FUNCTION "ROLL_PB13" : Void
{ S7_Optimized_Access := 'TRUE' }
VERSION : 0.1
VAR_TEMP
    r : Bool;
    a1 : Word;
    a2 : Word;
    activeDataBlock : Int;
    comparisonResults : Array[0..0] of Bool;
END_VAR
BEGIN
    #r := FALSE;
    #a1 := W#16#0000;
    #a2 := W#16#0000;
    #activeDataBlock := 0;
    // PB13, STEP 5 network 1
    #r := ((NOT "ROLL_State".M[58, 6]) AND ("ROLL_IO".Input[11, 1] OR "ROLL_IO".Input[11, 2] OR "ROLL_IO".Input[11, 3] OR "ROLL_IO".Input[11, 4] OR "ROLL_IO".Input[119, 6] OR "ROLL_IO".Input[119, 7] OR "ROLL_IO".Input[120, 0]) AND "ROLL_IO".Input[11, 6]);
    IF #r THEN "ROLL_State".M[58, 7] := TRUE; END_IF;
    #r := (((NOT "ROLL_IO".Input[11, 6]) AND ("ROLL_IO".Input[11, 1] OR "ROLL_IO".Input[11, 2] OR "ROLL_IO".Input[11, 3] OR "ROLL_IO".Input[11, 4] OR "ROLL_IO".Input[119, 6] OR "ROLL_IO".Input[119, 7] OR "ROLL_IO".Input[120, 0]) AND "ROLL_IO".Output[23, 0] AND "ROLL_State".M[58, 6]) OR "ROLL_IO".Input[11, 0]);
    IF #r THEN "ROLL_State".M[58, 7] := FALSE; END_IF;
    // PB13, STEP 5 network 2
    #r := "ROLL_IO".Input[11, 6];
    "ROLL_State".M[58, 6] := #r;
    // PB13, STEP 5 network 3
    #r := (((((NOT "ROLL_IO".Input[11, 0]) OR "ROLL_State".M[80, 7]) AND "ROLL_IO".Input[11, 6]) OR "ROLL_State".M[58, 7]) AND "ROLL_IO".Input[14, 0]);
    "ROLL_State".M[60, 0] := #r;
    // PB13, STEP 5 network 4
    #a2 := #a1;
    #a1 := W#16#2030;
    #r := ((NOT "ROLL_IO".Input[13, 3]) AND "ROLL_IO".Output[24, 0]);
    "ROLL_TimerOp"(Number := 110, Operation := 0, Signal := #r, Preset := #a1);
    // PB13, STEP 5 network 5
    #r := (((NOT "ROLL_State".M[111, 1]) AND (NOT "ROLL_State".M[111, 2]) AND (NOT "ROLL_State".M[111, 5]) AND "ROLL_IO".Input[0, 2] AND "ROLL_State".M[111, 0]) OR ((NOT "ROLL_State".M[61, 5]) AND "ROLL_IO".Input[0, 1] AND "ROLL_State".M[23, 2]) OR ("ROLL_IO".Input[12, 1] AND "ROLL_State".M[111, 5]));
    "ROLL_State".M[60, 1] := #r;
    // PB13, STEP 5 network 6
    #r := (((NOT "ROLL_IO".Input[12, 1]) AND "ROLL_State".M[111, 5]) OR ((NOT "ROLL_State".M[111, 0]) AND (NOT "ROLL_State".M[111, 2]) AND (NOT "ROLL_State".M[111, 5]) AND "ROLL_IO".Input[0, 2] AND "ROLL_State".M[111, 1]) OR ("ROLL_IO".Input[0, 1] AND "ROLL_State".M[23, 3]));
    "ROLL_State".M[60, 3] := #r;
    // PB13, STEP 5 network 7
    #r := (((NOT "ROLL_State".M[111, 0]) AND (NOT "ROLL_State".M[111, 1]) AND (NOT "ROLL_State".M[111, 5]) AND "ROLL_IO".Input[0, 2] AND "ROLL_State".M[111, 2]) OR ((NOT "ROLL_State".M[61, 5]) AND "ROLL_IO".Input[0, 1] AND "ROLL_State".M[0, 3]));
    "ROLL_State".M[60, 2] := #r;
    // PB13, STEP 5 network 8
    #a2 := #a1;
    #a1 := W#16#0005;
    #r := (NOT "ROLL_State".S5Timers[114].Q);
    "ROLL_TimerOp"(Number := 113, Operation := 0, Signal := #r, Preset := #a1);
    #a2 := #a1;
    #a1 := W#16#0005;
    #r := "ROLL_State".S5Timers[113].Q;
    "ROLL_TimerOp"(Number := 114, Operation := 1, Signal := #r, Preset := #a1);
    // PB13, STEP 5 network 9
    #activeDataBlock := 15;
    // PB13, STEP 5 network 10
    #a2 := #a1;
    #a1 := "ROLL_GetDW"(DbNumber := #activeDataBlock, Index := 116);
    #r := ((NOT "ROLL_State".S5Timers[117].Q) AND "ROLL_State".M[62, 4]);
    "ROLL_TimerOp"(Number := 116, Operation := 0, Signal := #r, Preset := #a1);
    #a2 := #a1;
    #a1 := "ROLL_GetDW"(DbNumber := #activeDataBlock, Index := 117);
    #r := "ROLL_State".S5Timers[116].Q;
    "ROLL_TimerOp"(Number := 117, Operation := 1, Signal := #r, Preset := #a1);
    // PB13, STEP 5 network 11
    #activeDataBlock := 19;
    // PB13, STEP 5 network 12
    #r := ("ROLL_IO".Output[24, 2] AND "ROLL_State".M[60, 4] AND "ROLL_State".S5Timers[114].Q);
    "ROLL_CounterOp"(Number := 1, Operation := 3, Signal := #r, Preset := #a1);
    #a2 := #a1;
    #a1 := "ROLL_GetDW"(DbNumber := #activeDataBlock, Index := 1);
    #r := ((((NOT "ROLL_IO".Input[13, 3]) AND (NOT ("ROLL_State".S5Counters[1].Value <> 0)) AND (NOT ("ROLL_State".S5Counters[2].Value <> 0))) OR "ROLL_IO".Input[13, 3] OR "ROLL_State".M[60, 5]) AND "ROLL_State".S5Timers[114].Q);
    "ROLL_CounterOp"(Number := 1, Operation := 0, Signal := #r, Preset := #a1);
    // PB13, STEP 5 network 13
    #r := ("ROLL_IO".Output[24, 0] AND "ROLL_State".M[60, 5] AND "ROLL_State".S5Timers[114].Q);
    "ROLL_CounterOp"(Number := 2, Operation := 3, Signal := #r, Preset := #a1);
    #a2 := #a1;
    #a1 := "ROLL_GetDW"(DbNumber := #activeDataBlock, Index := 2);
    #r := (("ROLL_IO".Input[13, 3] OR "ROLL_State".M[60, 4]) AND "ROLL_State".S5Timers[114].Q);
    "ROLL_CounterOp"(Number := 2, Operation := 0, Signal := #r, Preset := #a1);
    // PB13, STEP 5 network 14
    #r := ((NOT "ROLL_IO".Input[13, 3]) AND "ROLL_IO".Output[24, 2] AND "ROLL_State".M[60, 6]);
    IF #r THEN "ROLL_State".M[60, 4] := TRUE; END_IF;
    #r := "ROLL_IO".Input[13, 3];
    IF #r THEN "ROLL_State".M[60, 4] := FALSE; END_IF;
    // PB13, STEP 5 network 15
    #r := ((NOT "ROLL_IO".Input[13, 3]) AND "ROLL_IO".Output[24, 0] AND "ROLL_State".M[60, 6]);
    IF #r THEN "ROLL_State".M[60, 5] := TRUE; END_IF;
    #r := "ROLL_IO".Input[13, 3];
    IF #r THEN "ROLL_State".M[60, 5] := FALSE; END_IF;
    // PB13, STEP 5 network 16
    #r := "ROLL_IO".Input[13, 3];
    IF #r THEN "ROLL_State".M[60, 6] := TRUE; END_IF;
    #r := ("ROLL_State".M[60, 4] OR "ROLL_State".M[60, 5]);
    IF #r THEN "ROLL_State".M[60, 6] := FALSE; END_IF;
    // PB13, STEP 5 network 17
    #r := ((NOT ("ROLL_State".S5Counters[2].Value <> 0)) AND "ROLL_State".M[62, 6]);
    IF #r THEN "ROLL_State".M[60, 7] := TRUE; END_IF;
    #r := (NOT "ROLL_State".M[62, 6]);
    IF #r THEN "ROLL_State".M[60, 7] := FALSE; END_IF;
    // PB13, STEP 5 network 18
    #r := ((NOT "ROLL_IO".Input[13, 3]) AND (NOT ("ROLL_State".S5Counters[1].Value <> 0)) AND "ROLL_State".M[61, 1]);
    IF #r THEN "ROLL_State".M[61, 0] := TRUE; END_IF;
    #r := (NOT "ROLL_State".M[62, 6]);
    IF #r THEN "ROLL_State".M[61, 0] := FALSE; END_IF;
    // PB13, STEP 5 network 19
    #r := ("ROLL_State".S5Counters[1].Value <> 0);
    "ROLL_State".M[61, 1] := #r;
    // PB13, STEP 5 network 20
    #r := (("ROLL_State".M[60, 7] OR "ROLL_State".M[62, 6]) AND "ROLL_State".M[61, 0]);
    "ROLL_State".M[61, 2] := #r;
    // PB13, STEP 5 network 21
    #r := ((NOT "ROLL_State".M[61, 6]) AND "ROLL_State".M[60, 1] AND "ROLL_State".M[61, 7]);
    IF #r THEN "ROLL_State".M[61, 3] := TRUE; END_IF;
    #r := (NOT "ROLL_State".M[61, 7]);
    IF #r THEN "ROLL_State".M[61, 3] := FALSE; END_IF;
    // PB13, STEP 5 network 22
    #r := ((NOT "ROLL_State".M[61, 6]) AND "ROLL_State".M[60, 2] AND "ROLL_State".M[61, 7]);
    IF #r THEN "ROLL_State".M[61, 4] := TRUE; END_IF;
    #r := (NOT "ROLL_State".M[61, 7]);
    IF #r THEN "ROLL_State".M[61, 4] := FALSE; END_IF;
    // PB13, STEP 5 network 23
    #r := ((NOT "ROLL_State".M[61, 6]) AND "ROLL_State".M[60, 3] AND "ROLL_State".M[61, 7]);
    IF #r THEN "ROLL_State".M[61, 5] := TRUE; END_IF;
    #r := (NOT "ROLL_State".M[61, 7]);
    IF #r THEN "ROLL_State".M[61, 5] := FALSE; END_IF;
    // PB13, STEP 5 network 24
    #r := "ROLL_State".M[61, 7];
    "ROLL_State".M[61, 6] := #r;
    // PB13, STEP 5 network 25
    #r := (((NOT "ROLL_State".M[111, 5]) AND "ROLL_State".M[37, 3]) OR ((((NOT "ROLL_IO".Input[12, 1]) AND ("ROLL_State".M[41, 0] OR "ROLL_State".M[42, 4] OR "ROLL_State".M[44, 0])) OR (("ROLL_State".M[40, 5] OR "ROLL_State".M[42, 1] OR "ROLL_State".M[43, 5]) AND "ROLL_IO".Input[12, 1])) AND "ROLL_State".M[111, 5]));
    IF #r THEN "ROLL_State".M[61, 7] := TRUE; END_IF;
    #r := (((NOT "ROLL_IO".Input[12, 5]) AND "ROLL_IO".Input[11, 0] AND "ROLL_State".M[190, 5] AND "ROLL_State".M[20, 1]) OR (("ROLL_State".M[42, 0] OR "ROLL_State".M[43, 4] OR "ROLL_State".M[58, 5]) AND "ROLL_State".M[111, 5]) OR "ROLL_State".M[53, 6]);
    IF #r THEN "ROLL_State".M[61, 7] := FALSE; END_IF;
    // PB13, STEP 5 network 26
    #r := ((NOT "ROLL_IO".Input[11, 0]) AND (((NOT "ROLL_IO".Input[12, 1]) AND "ROLL_IO".Output[23, 5]) OR ("ROLL_IO".Output[23, 4] AND "ROLL_IO".Input[12, 1])) AND ("ROLL_State".M[61, 3] OR "ROLL_State".M[61, 4] OR "ROLL_State".M[61, 5]));
    IF #r THEN "ROLL_State".M[62, 0] := TRUE; END_IF;
    #r := ((("ROLL_State".M[41, 3] OR "ROLL_State".M[42, 7] OR "ROLL_State".M[44, 3] OR "ROLL_State".M[46, 0] OR "ROLL_State".M[47, 3] OR "ROLL_State".M[48, 7] OR "ROLL_State".M[50, 3] OR "ROLL_State".M[51, 5]) AND "ROLL_IO".Input[13, 3] AND "ROLL_State".S5Timers[114].Q) OR (NOT "ROLL_State".M[31, 5]) OR (NOT "ROLL_State".M[61, 7]));
    IF #r THEN "ROLL_State".M[62, 0] := FALSE; END_IF;
    // PB13, STEP 5 network 27
    #r := (((NOT "ROLL_IO".Input[11, 0]) AND ((("ROLL_IO".Input[11, 1] OR "ROLL_IO".Input[11, 2] OR "ROLL_IO".Input[11, 3] OR "ROLL_IO".Input[11, 4] OR "ROLL_IO".Input[119, 6] OR "ROLL_IO".Input[119, 7] OR "ROLL_IO".Input[120, 0]) AND ("ROLL_State".M[80, 6] OR "ROLL_State".M[80, 7])) OR ("ROLL_State".M[60, 0] AND "ROLL_State".M[80, 7]))) OR ("ROLL_IO".Input[11, 0] AND "ROLL_IO".Input[11, 6] AND "ROLL_State".M[80, 7]));
    "ROLL_State".M[62, 1] := #r;
    // PB13, STEP 5 network 28
    #r := (("ROLL_State".M[0, 3] AND "ROLL_State".M[45, 6]) OR "ROLL_State".M[41, 1] OR "ROLL_State".M[42, 5] OR "ROLL_State".M[44, 1] OR "ROLL_State".M[47, 1] OR "ROLL_State".M[48, 5] OR "ROLL_State".M[50, 1]);
    "ROLL_State".M[63, 5] := #r;
    // PB13, STEP 5 network 29
    #r := (((((NOT "ROLL_State".M[60, 1]) AND (NOT "ROLL_State".M[60, 2]) AND (NOT "ROLL_State".M[60, 3]) AND (NOT "ROLL_State".M[63, 1]) AND "ROLL_State".M[74, 0]) OR ((NOT "ROLL_State".M[60, 1]) AND (NOT "ROLL_State".M[60, 2]) AND "ROLL_State".M[60, 3])) AND ("ROLL_State".M[20, 1] OR "ROLL_State".M[20, 2] OR "ROLL_State".M[23, 3]) AND "ROLL_IO".Input[0, 1]) OR ((((NOT "ROLL_State".M[61, 3]) AND (NOT "ROLL_State".M[61, 4]) AND (NOT "ROLL_State".M[61, 5]) AND "ROLL_State".M[62, 6]) OR ((NOT "ROLL_State".M[61, 3]) AND (NOT "ROLL_State".M[61, 4]) AND "ROLL_State".M[61, 5])) AND "ROLL_IO".Input[0, 2]));
    "ROLL_State".M[62, 2] := #r;
    // PB13, STEP 5 network 30
    #r := (((NOT "ROLL_State".M[60, 2]) AND (NOT "ROLL_State".M[60, 3]) AND ("ROLL_State".M[20, 1] OR "ROLL_State".M[23, 2]) AND "ROLL_IO".Input[0, 1] AND "ROLL_State".M[60, 1]) OR ((NOT "ROLL_State".M[61, 4]) AND (NOT "ROLL_State".M[61, 5]) AND (NOT "ROLL_State".M[63, 5]) AND "ROLL_IO".Input[0, 2] AND "ROLL_State".M[61, 3]));
    "ROLL_State".M[62, 3] := #r;
    // PB13, STEP 5 network 31
    #r := (((NOT "ROLL_State".M[60, 1]) AND (NOT "ROLL_State".M[60, 3]) AND ("ROLL_State".M[0, 3] OR "ROLL_State".M[20, 1]) AND "ROLL_IO".Input[0, 1] AND "ROLL_State".M[60, 2]) OR ((((NOT "ROLL_State".M[61, 3]) AND (NOT "ROLL_State".M[61, 5]) AND "ROLL_State".M[61, 4]) OR ("ROLL_State".M[61, 3] AND "ROLL_State".M[63, 5])) AND "ROLL_IO".Input[0, 2]));
    "ROLL_State".M[62, 4] := #r;
    // PB13, STEP 5 network 32
    #r := ((((NOT "ROLL_State".M[190, 5]) AND ("ROLL_State".M[0, 3] OR "ROLL_State".M[23, 2] OR "ROLL_State".M[23, 3]) AND ("ROLL_State".M[60, 1] OR "ROLL_State".M[60, 2] OR "ROLL_State".M[60, 3]) AND "ROLL_IO".Input[0, 1] AND "ROLL_State".M[190, 6] AND "ROLL_State".M[62, 1]) OR ("ROLL_IO".Input[0, 2] AND "ROLL_State".M[31, 5] AND "ROLL_State".M[62, 0])) AND ("ROLL_State".M[62, 5] OR "ROLL_State".S5Timers[114].Q) AND "ROLL_State".M[60, 0]);
    "ROLL_State".M[62, 5] := #r;
    // PB13, STEP 5 network 33
    #r := ((NOT "ROLL_State".M[63, 1]) AND (((NOT "ROLL_State".M[62, 0]) AND "ROLL_IO".Input[0, 2] AND "ROLL_State".M[31, 5]) OR ((((NOT "ROLL_State".M[190, 6]) AND ("ROLL_State".M[0, 3] OR "ROLL_State".M[20, 2] OR "ROLL_State".M[23, 2] OR "ROLL_State".M[23, 3]) AND "ROLL_State".M[190, 5]) OR "ROLL_State".M[74, 0]) AND "ROLL_IO".Input[0, 1] AND "ROLL_State".M[62, 1])) AND ("ROLL_State".M[62, 6] OR "ROLL_State".S5Timers[114].Q) AND "ROLL_State".M[60, 0]);
    "ROLL_State".M[62, 6] := #r;
    // PB13, STEP 5 network 34
    #r := ((((NOT "ROLL_State".M[61, 2]) AND (NOT "ROLL_State".M[63, 1]) AND "ROLL_State".M[62, 6]) OR "ROLL_State".M[62, 5]) AND (((NOT "ROLL_State".M[62, 2]) AND (NOT "ROLL_State".M[62, 4]) AND (NOT "ROLL_State".M[62, 6]) AND "ROLL_State".M[62, 3]) OR ((NOT "ROLL_State".M[62, 6]) AND ("ROLL_IO".Input[13, 3] OR "ROLL_State".S5Timers[117].Q) AND "ROLL_State".M[62, 4]) OR (((NOT "ROLL_State".M[62, 4]) OR "ROLL_State".M[62, 6]) AND ("ROLL_State".S5Counters[1].Value <> 0))) AND ("ROLL_State".M[62, 2] OR "ROLL_State".M[62, 3] OR "ROLL_State".M[62, 4]));
    "ROLL_State".M[62, 7] := #r;
    // PB13, STEP 5 network 35
    #r := ((NOT "ROLL_IO".Output[24, 0]) AND (NOT "ROLL_State".M[5, 1]) AND (NOT "ROLL_State".M[63, 4]) AND ((NOT "ROLL_State".S5Timers[115].Q) OR "ROLL_IO".Output[24, 2]) AND "ROLL_IO".Input[13, 5] AND "ROLL_State".M[29, 0] AND "ROLL_State".M[60, 0] AND "ROLL_State".M[62, 7]);
    "ROLL_IO".Output[24, 2] := #r;
    // PB13, STEP 5 network 36
    #r := ((((NOT "ROLL_State".M[62, 2]) AND (NOT "ROLL_State".M[62, 6])) OR ("ROLL_State".S5Counters[2].Value <> 0)) AND (((NOT "ROLL_State".M[63, 1]) AND "ROLL_State".M[62, 6]) OR "ROLL_State".M[62, 5]) AND ((NOT "ROLL_State".M[62, 4]) OR (NOT "ROLL_State".M[62, 5])));
    "ROLL_State".M[63, 0] := #r;
    // PB13, STEP 5 network 37
    #r := ((NOT "ROLL_IO".Output[24, 2]) AND (NOT "ROLL_State".M[5, 1]) AND (NOT "ROLL_State".M[63, 4]) AND ((NOT "ROLL_State".S5Timers[115].Q) OR "ROLL_IO".Output[24, 0]) AND "ROLL_IO".Input[13, 5] AND "ROLL_State".M[29, 0] AND "ROLL_State".M[60, 0] AND "ROLL_State".M[63, 0]);
    "ROLL_IO".Output[24, 0] := #r;
    // PB13, STEP 5 network 38
    #r := ((NOT "ROLL_IO".Output[24, 5]) AND "ROLL_IO".Output[24, 0] AND "ROLL_IO".Input[13, 3]);
    "ROLL_IO".Output[24, 1] := #r;
    // PB13, STEP 5 network 39
    #r := ("ROLL_IO".Output[24, 0] OR "ROLL_IO".Output[24, 2] OR "ROLL_State".M[63, 6]);
    "ROLL_State".M[240, 0] := #r;
    // PB13, STEP 5 network 40
    #r := ((NOT "ROLL_IO".Input[12, 5]) AND (("ROLL_State".M[190, 5] AND "ROLL_State".M[23, 0]) OR "ROLL_State".M[52, 2]) AND "ROLL_IO".Input[11, 0] AND "ROLL_IO".Input[11, 6]);
    IF #r THEN "ROLL_State".M[63, 6] := TRUE; END_IF;
    #r := (("ROLL_IO".Input[12, 1] OR "ROLL_IO".Input[12, 5]) AND "ROLL_IO".Input[11, 0] AND "ROLL_IO".Input[11, 6] AND "ROLL_IO".Input[12, 7]);
    IF #r THEN "ROLL_State".M[63, 6] := FALSE; END_IF;
    // PB13, STEP 5 network 41
    #r := ((((NOT "ROLL_State".M[63, 7]) AND "ROLL_IO".Output[24, 0] AND "ROLL_State".S5Timers[111].Q) OR ("ROLL_IO".Input[11, 0] AND "ROLL_State".M[80, 6]) OR (NOT "ROLL_State".S5Timers[11].Q)) AND "ROLL_IO".Input[13, 3]);
    IF #r THEN "ROLL_State".M[63, 1] := TRUE; END_IF;
    #r := (((NOT "ROLL_IO".Input[13, 3]) AND "ROLL_IO".Input[3, 0] AND "ROLL_State".S5Timers[11].Q) OR "ROLL_IO".Output[24, 2]);
    IF #r THEN "ROLL_State".M[63, 1] := FALSE; END_IF;
    // PB13, STEP 5 network 42
    #a2 := #a1;
    #a1 := W#16#1030;
    #r := ("ROLL_IO".Output[24, 0] AND "ROLL_IO".Input[13, 3] AND "ROLL_State".M[29, 0] AND "ROLL_State".M[61, 2]);
    "ROLL_TimerOp"(Number := 111, Operation := 0, Signal := #r, Preset := #a1);
    // PB13, STEP 5 network 43
    #r := (((NOT "ROLL_IO".Input[13, 3]) AND "ROLL_IO".Input[0, 1] AND "ROLL_State".M[0, 3] AND "ROLL_State".M[190, 6]) OR ((((NOT "ROLL_State".M[61, 2]) AND "ROLL_State".M[62, 6]) OR "ROLL_State".M[62, 5]) AND ("ROLL_State".M[62, 2] OR "ROLL_State".M[62, 3] OR "ROLL_State".M[62, 4])) OR ("ROLL_IO".Input[13, 3] AND "ROLL_State".M[63, 7]));
    "ROLL_State".M[63, 7] := #r;
    "ROLL_IO".Output[24, 5] := #r;
    // PB13, STEP 5 network 44
    #r := ("ROLL_IO".Output[24, 0] OR "ROLL_IO".Output[24, 2]);
    "ROLL_IO".Output[24, 4] := #r;
    // PB13, STEP 5 network 45
    #r := ("ROLL_State".M[41, 1] OR "ROLL_State".M[42, 5] OR "ROLL_State".M[44, 1] OR "ROLL_State".M[45, 6] OR "ROLL_State".M[47, 1] OR "ROLL_State".M[48, 5] OR "ROLL_State".M[50, 1]);
    "ROLL_State".M[240, 0] := #r;
    // PB13, STEP 5 network 46
    #r := "ROLL_State".M[111, 1];
    "ROLL_State".M[240, 1] := #r;
    // PB13, STEP 5 network 47
    "ROLL_FB69"();
    // PB13, STEP 5 network 48
    #a2 := #a1;
    #a1 := "ROLL_GetM"(FirstByte := 240, Width := 16);
    #r := ("ROLL_IO".Output[24, 0] OR "ROLL_IO".Output[24, 2]);
    "ROLL_TimerOp"(Number := 115, Operation := 1, Signal := #r, Preset := #a1);
    // PB13, STEP 5 network 49
    #r := ((("ROLL_IO".Output[24, 0] AND "ROLL_State".M[60, 5]) OR ("ROLL_IO".Output[24, 2] AND "ROLL_State".M[60, 4])) AND "ROLL_State".S5Timers[114].Q);
    "ROLL_CounterOp"(Number := 3, Operation := 3, Signal := #r, Preset := #a1);
    #r := ((((NOT "ROLL_State".M[60, 4]) AND (NOT "ROLL_State".M[60, 5]) AND ("ROLL_IO".Output[24, 0] OR "ROLL_IO".Output[24, 2])) OR ("ROLL_IO".Output[24, 0] AND "ROLL_State".M[60, 4]) OR ("ROLL_IO".Output[24, 2] AND "ROLL_State".M[60, 5])) AND "ROLL_State".S5Timers[114].Q);
    "ROLL_CounterOp"(Number := 3, Operation := 2, Signal := #r, Preset := #a1);
    #a2 := #a1;
    #a1 := W#16#0500;
    #r := (("ROLL_IO".Input[13, 3] AND "ROLL_State".S5Timers[114].Q) OR ("ROLL_State".M[3, 1] AND "ROLL_State".M[63, 2]));
    "ROLL_CounterOp"(Number := 3, Operation := 0, Signal := #r, Preset := #a1);
    // PB13, STEP 5 network 50
    #a2 := #a1;
    #a1 := INT_TO_WORD("ROLL_State".S5Counters[3].Value);
    #a2 := #a1;
    #a1 := W#16#0208;
    #comparisonResults[0] := (WORD_TO_INT(#a2) > WORD_TO_INT(#a1));
    #r := #comparisonResults[0];
    "ROLL_State".M[63, 2] := #r;
    // PB13, STEP 5 network 51
    #a2 := #a1;
    #a1 := W#16#1060;
    #r := ((("ROLL_IO".Output[24, 0] AND "ROLL_State".M[63, 7]) OR "ROLL_IO".Output[24, 2]) AND "ROLL_IO".Input[13, 3]);
    "ROLL_TimerOp"(Number := 112, Operation := 0, Signal := #r, Preset := #a1);
    // PB13, STEP 5 network 52
    #r := ((NOT ("ROLL_State".S5Counters[2].Value <> 0)) AND "ROLL_State".M[61, 2] AND "ROLL_State".M[62, 6] AND ("ROLL_State".S5Counters[1].Value <> 0));
    "ROLL_State".M[63, 3] := #r;
    // PB13, STEP 5 network 53
    #r := (((NOT "ROLL_IO".Input[0, 4]) AND "ROLL_IO".Input[0, 2] AND "ROLL_State".M[63, 4]) OR "ROLL_State".M[11, 0] OR "ROLL_State".M[11, 1] OR "ROLL_State".M[11, 2] OR "ROLL_State".M[11, 3]);
    "ROLL_State".M[63, 4] := #r;
    // PB13, STEP 5 network 54
    RETURN;
END_FUNCTION

FUNCTION "ROLL_PB14" : Void
{ S7_Optimized_Access := 'TRUE' }
VERSION : 0.1
VAR_TEMP
    r : Bool;
    a1 : Word;
    a2 : Word;
    activeDataBlock : Int;
    comparisonResults : Array[0..0] of Bool;
END_VAR
BEGIN
    #r := FALSE;
    #a1 := W#16#0000;
    #a2 := W#16#0000;
    #activeDataBlock := 0;
    // PB14, STEP 5 network 1
    #activeDataBlock := 15;
    // PB14, STEP 5 network 2
    #r := ((NOT "ROLL_State".M[37, 5]) AND (NOT "ROLL_State".M[53, 2]) AND (NOT "ROLL_State".M[53, 3]) AND (((NOT "ROLL_State".S5Timers[21].Q) AND "ROLL_IO".Input[123, 4] AND "ROLL_State".M[31, 4]) OR ("ROLL_State".M[70, 4] AND "ROLL_State".S5Timers[45].Q) OR "ROLL_State".M[37, 7] OR "ROLL_State".M[53, 4] OR "ROLL_State".M[70, 7]) AND ((NOT "ROLL_State".S5Timers[95].Q) OR "ROLL_State".M[53, 4]) AND "ROLL_State".M[31, 5] AND "ROLL_State".M[35, 2]);
    "ROLL_State".M[64, 0] := #r;
    // PB14, STEP 5 network 3
    #r := (((NOT "ROLL_State".M[31, 4]) AND (NOT "ROLL_State".M[31, 5]) AND "ROLL_IO".Input[125, 4]) OR ((((NOT "ROLL_IO".Output[113, 4]) AND "ROLL_IO".Output[113, 5] AND "ROLL_State".M[72, 1]) OR "ROLL_State".M[53, 4]) AND "ROLL_State".M[31, 5] AND "ROLL_State".M[35, 2]));
    "ROLL_State".M[64, 1] := #r;
    // PB14, STEP 5 network 4
    #r := ("ROLL_IO".Input[123, 4] AND "ROLL_State".S5Timers[20].Q);
    IF #r THEN "ROLL_State".M[64, 4] := TRUE; END_IF;
    #r := (((NOT "ROLL_IO".Output[113, 3]) AND (NOT "ROLL_IO".Input[123, 4])) OR (NOT "ROLL_State".M[31, 5]));
    IF #r THEN "ROLL_State".M[64, 4] := FALSE; END_IF;
    // PB14, STEP 5 network 5
    #r := "ROLL_State".M[37, 5];
    IF #r THEN "ROLL_State".M[64, 5] := TRUE; END_IF;
    #r := ((NOT "ROLL_State".M[31, 5]) OR "ROLL_State".M[39, 5]);
    IF #r THEN "ROLL_State".M[64, 5] := FALSE; END_IF;
    // PB14, STEP 5 network 6
    #r := ((("ROLL_State".M[40, 2] OR "ROLL_State".M[44, 7] OR "ROLL_State".M[50, 6]) AND "ROLL_State".M[63, 1]) OR "ROLL_State".M[41, 6] OR "ROLL_State".M[43, 2] OR "ROLL_State".M[44, 7] OR "ROLL_State".M[46, 2] OR "ROLL_State".M[47, 6] OR "ROLL_State".M[49, 2]);
    "ROLL_State".M[65, 0] := #r;
    // PB14, STEP 5 network 7
    #r := ("ROLL_IO".Input[12, 5] AND "ROLL_IO".Input[12, 7] AND "ROLL_State".M[52, 0] AND "ROLL_State".M[63, 1]);
    "ROLL_State".M[65, 5] := #r;
    // PB14, STEP 5 network 8
    #r := (((NOT "ROLL_IO".Input[11, 0]) AND "ROLL_State".M[52, 0]) OR ((NOT "ROLL_IO".Input[11, 1]) AND "ROLL_State".M[40, 2]) OR ((NOT "ROLL_IO".Input[11, 2]) AND "ROLL_State".M[41, 6]) OR ((NOT "ROLL_IO".Input[11, 3]) AND "ROLL_State".M[43, 2]) OR ((NOT "ROLL_IO".Input[11, 4]) AND "ROLL_State".M[44, 7]) OR ((NOT "ROLL_IO".Input[119, 6]) AND "ROLL_State".M[46, 2]) OR ((NOT "ROLL_IO".Input[119, 7]) AND "ROLL_State".M[47, 6]) OR ((NOT "ROLL_IO".Input[120, 0]) AND "ROLL_State".M[49, 2]) OR ((NOT "ROLL_IO".Input[120, 1]) AND "ROLL_State".M[50, 6]));
    "ROLL_State".M[65, 6] := #r;
    // PB14, STEP 5 network 9
    #r := (("ROLL_IO".Input[11, 0] AND "ROLL_State".M[40, 0]) OR ("ROLL_IO".Input[11, 1] AND "ROLL_State".M[41, 0]) OR ("ROLL_IO".Input[11, 2] AND "ROLL_State".M[42, 4]) OR ("ROLL_IO".Input[11, 3] AND "ROLL_State".M[44, 0]) OR ("ROLL_IO".Input[11, 4] AND "ROLL_State".M[45, 5]) OR ("ROLL_IO".Input[119, 6] AND "ROLL_State".M[47, 0]) OR ("ROLL_IO".Input[119, 7] AND "ROLL_State".M[48, 4]) OR ("ROLL_IO".Input[120, 0] AND "ROLL_State".M[50, 0]) OR ("ROLL_IO".Input[120, 1] AND "ROLL_State".M[51, 3]));
    "ROLL_State".M[66, 2] := #r;
    // PB14, STEP 5 network 10
    #r := (("ROLL_State".M[66, 2] OR "ROLL_State".M[68, 2]) AND "ROLL_IO".Input[11, 6]);
    "ROLL_State".M[66, 4] := #r;
    // PB14, STEP 5 network 11
    #r := (("ROLL_IO".Input[11, 1] AND "ROLL_State".M[40, 4]) OR ("ROLL_IO".Input[11, 2] AND "ROLL_State".M[42, 0]) OR ("ROLL_IO".Input[11, 3] AND "ROLL_State".M[43, 4]) OR ("ROLL_IO".Input[11, 4] AND "ROLL_State".M[45, 1]) OR ("ROLL_IO".Input[119, 6] AND "ROLL_State".M[46, 4]) OR ("ROLL_IO".Input[119, 7] AND "ROLL_State".M[48, 0]) OR ("ROLL_IO".Input[120, 0] AND "ROLL_State".M[49, 4]) OR ("ROLL_IO".Input[120, 1] AND "ROLL_State".M[51, 0]));
    "ROLL_State".M[66, 5] := #r;
    // PB14, STEP 5 network 12
    #r := (((NOT "ROLL_IO".Input[12, 1]) OR (NOT "ROLL_IO".Input[12, 7])) AND "ROLL_IO".Input[11, 0] AND "ROLL_State".M[52, 2]);
    "ROLL_State".M[66, 6] := #r;
    // PB14, STEP 5 network 13
    #r := (("ROLL_State".M[66, 5] OR "ROLL_State".M[66, 6] OR "ROLL_State".M[68, 3]) AND "ROLL_IO".Input[11, 6]);
    "ROLL_State".M[66, 7] := #r;
    // PB14, STEP 5 network 14
    #r := ((NOT "ROLL_IO".Output[113, 3]) AND (NOT "ROLL_State".M[9, 3]) AND "ROLL_IO".Input[124, 5] AND "ROLL_State".M[39, 6]);
    "ROLL_State".M[67, 0] := #r;
    // PB14, STEP 5 network 15
    #r := ((NOT "ROLL_IO".Output[113, 3]) AND (NOT "ROLL_State".M[9, 3]) AND "ROLL_IO".Input[124, 5] AND "ROLL_State".M[53, 0]);
    "ROLL_State".M[67, 1] := #r;
    // PB14, STEP 5 network 16
    #r := ((NOT "ROLL_IO".Input[124, 5]) AND "ROLL_IO".Input[124, 1] AND "ROLL_State".M[39, 4]);
    "ROLL_State".M[67, 5] := #r;
    // PB14, STEP 5 network 17
    #r := ((NOT "ROLL_IO".Input[124, 4]) AND "ROLL_IO".Input[124, 1] AND "ROLL_State".M[53, 2]);
    "ROLL_State".M[67, 6] := #r;
    // PB14, STEP 5 network 18
    #r := ((("ROLL_IO".Input[5, 1] AND "ROLL_State".M[40, 5]) OR ("ROLL_State".M[0, 3] AND "ROLL_State".M[45, 2]) OR "ROLL_State".M[42, 1] OR "ROLL_State".M[43, 5] OR "ROLL_State".M[46, 5] OR "ROLL_State".M[48, 1] OR "ROLL_State".M[49, 5]) AND "ROLL_State".M[111, 3]);
    "ROLL_State".M[68, 0] := #r;
    // PB14, STEP 5 network 19
    #r := ((NOT "ROLL_State".S5Timers[25].Q) AND (("ROLL_IO".Input[12, 1] AND "ROLL_IO".Input[12, 7]) OR "ROLL_State".M[68, 2]) AND ("ROLL_State".M[68, 2] OR "ROLL_State".S5Timers[24].Q) AND "ROLL_State".M[68, 0]);
    "ROLL_State".M[68, 2] := #r;
    // PB14, STEP 5 network 20
    #r := (((NOT "ROLL_IO".Input[12, 1]) OR (NOT "ROLL_IO".Input[12, 7])) AND ("ROLL_State".M[68, 3] OR "ROLL_State".S5Timers[24].Q) AND "ROLL_State".M[68, 0]);
    "ROLL_State".M[68, 3] := #r;
    // PB14, STEP 5 network 21
    #a2 := #a1;
    #a1 := "ROLL_GetDW"(DbNumber := #activeDataBlock, Index := 24);
    #r := ((NOT "ROLL_State".M[68, 2]) AND (NOT "ROLL_State".M[68, 3]));
    "ROLL_TimerOp"(Number := 24, Operation := 0, Signal := #r, Preset := #a1);
    // PB14, STEP 5 network 22
    #a2 := #a1;
    #a1 := "ROLL_GetDW"(DbNumber := #activeDataBlock, Index := 25);
    #r := "ROLL_State".M[68, 2];
    "ROLL_TimerOp"(Number := 25, Operation := 0, Signal := #r, Preset := #a1);
    // PB14, STEP 5 network 23
    RETURN;
END_FUNCTION

FUNCTION "ROLL_PB15" : Void
{ S7_Optimized_Access := 'TRUE' }
VERSION : 0.1
VAR_TEMP
    r : Bool;
    a1 : Word;
    a2 : Word;
    activeDataBlock : Int;
    comparisonResults : Array[0..0] of Bool;
END_VAR
BEGIN
    #r := FALSE;
    #a1 := W#16#0000;
    #a2 := W#16#0000;
    #activeDataBlock := 0;
    // PB15, STEP 5 network 1
    #r := ((NOT "ROLL_IO".Output[113, 2]) AND "ROLL_IO".Output[113, 3] AND "ROLL_IO".Input[123, 4]);
    IF #r THEN "ROLL_State".M[70, 2] := TRUE; END_IF;
    #r := (((NOT "ROLL_IO".Input[123, 4]) AND "ROLL_IO".Input[123, 5]) OR "ROLL_State".M[73, 7]);
    IF #r THEN "ROLL_State".M[70, 2] := FALSE; END_IF;
    // PB15, STEP 5 network 2
    #r := ((((NOT "ROLL_State".M[20, 2]) AND "ROLL_IO".Input[123, 6] AND "ROLL_State".M[74, 0]) OR "ROLL_State".M[71, 0]) AND "ROLL_IO".Output[113, 2] AND "ROLL_IO".Input[124, 1] AND "ROLL_IO".Input[124, 4]);
    IF #r THEN "ROLL_State".M[70, 3] := TRUE; END_IF;
    #r := (((NOT "ROLL_IO".Input[123, 5]) AND (NOT "ROLL_IO".Input[123, 6])) OR "ROLL_State".M[73, 7]);
    IF #r THEN "ROLL_State".M[70, 3] := FALSE; END_IF;
    // PB15, STEP 5 network 3
    #r := ((NOT "ROLL_State".M[16, 0]) AND (NOT "ROLL_State".M[16, 1]) AND (NOT "ROLL_State".M[16, 4]) AND (NOT "ROLL_State".M[71, 1]) AND "ROLL_IO".Input[123, 1] AND "ROLL_State".M[191, 4] AND "ROLL_State".M[31, 4] AND "ROLL_State".S5Timers[45].Q);
    IF #r THEN "ROLL_State".M[70, 4] := TRUE; END_IF;
    #r := ((NOT "ROLL_IO".Input[123, 1]) OR "ROLL_State".M[73, 7]);
    IF #r THEN "ROLL_State".M[70, 4] := FALSE; END_IF;
    // PB15, STEP 5 network 4
    #r := "ROLL_IO".Input[123, 6];
    IF #r THEN "ROLL_State".M[70, 5] := TRUE; END_IF;
    #r := ("ROLL_IO".Input[125, 0] OR "ROLL_State".M[73, 7]);
    IF #r THEN "ROLL_State".M[70, 5] := FALSE; END_IF;
    // PB15, STEP 5 network 5
    #r := ((NOT "ROLL_IO".Input[125, 1]) AND "ROLL_IO".Output[113, 4] AND "ROLL_IO".Input[125, 0]);
    IF #r THEN "ROLL_State".M[70, 6] := TRUE; END_IF;
    #r := (("ROLL_IO".Output[113, 5] AND "ROLL_IO".Input[125, 1]) OR "ROLL_State".M[73, 7]);
    IF #r THEN "ROLL_State".M[70, 6] := FALSE; END_IF;
    // PB15, STEP 5 network 6
    #r := ((NOT "ROLL_State".M[71, 1]) AND "ROLL_IO".Input[123, 1] AND "ROLL_State".S5Timers[45].Q);
    IF #r THEN "ROLL_State".M[70, 7] := TRUE; END_IF;
    #r := ("ROLL_IO".Input[123, 4] OR "ROLL_State".M[73, 7]);
    IF #r THEN "ROLL_State".M[70, 7] := FALSE; END_IF;
    // PB15, STEP 5 network 7
    #r := ("ROLL_IO".Output[113, 3] AND "ROLL_IO".Input[123, 5]);
    IF #r THEN "ROLL_State".M[71, 0] := TRUE; END_IF;
    #r := ("ROLL_State".M[70, 3] OR "ROLL_State".M[73, 7]);
    IF #r THEN "ROLL_State".M[71, 0] := FALSE; END_IF;
    // PB15, STEP 5 network 8
    #r := ((NOT "ROLL_State".M[190, 6]) AND (NOT "ROLL_State".M[28, 4]) AND ("ROLL_State".M[20, 1] OR "ROLL_State".M[20, 2]) AND "ROLL_IO".Input[0, 1] AND "ROLL_State".M[190, 5]);
    "ROLL_State".M[74, 0] := #r;
    // PB15, STEP 5 network 9
    RETURN;
END_FUNCTION

FUNCTION "ROLL_PB16" : Void
{ S7_Optimized_Access := 'TRUE' }
VERSION : 0.1
VAR_TEMP
    r : Bool;
    a1 : Word;
    a2 : Word;
    activeDataBlock : Int;
    comparisonResults : Array[0..0] of Bool;
END_VAR
BEGIN
    #r := FALSE;
    #a1 := W#16#0000;
    #a2 := W#16#0000;
    #activeDataBlock := 0;
    // PB16, STEP 5 network 1
    #r := ("ROLL_IO".Input[0, 1] AND "ROLL_State".M[190, 5] AND "ROLL_State".M[190, 6] AND "ROLL_State".M[27, 7]);
    "ROLL_State".M[73, 7] := #r;
    // PB16, STEP 5 network 2
    #r := (("ROLL_State".M[20, 3] OR "ROLL_State".M[20, 5]) AND "ROLL_IO".Input[124, 1] AND "ROLL_IO".Input[124, 4]);
    "ROLL_State".M[74, 2] := #r;
    // PB16, STEP 5 network 3
    #r := (((NOT "ROLL_State".M[190, 5]) AND "ROLL_State".M[190, 6] AND "ROLL_State".M[74, 2]) OR (("ROLL_State".M[70, 2] OR "ROLL_State".M[70, 3]) AND "ROLL_State".M[74, 0]));
    "ROLL_State".M[74, 1] := #r;
    // PB16, STEP 5 network 4
    #r := (("ROLL_State".M[20, 4] OR "ROLL_State".M[20, 5]) AND "ROLL_IO".Input[0, 1] AND "ROLL_State".M[190, 6]);
    "ROLL_State".M[74, 4] := #r;
    // PB16, STEP 5 network 5
    #r := ((NOT "ROLL_IO".Output[113, 3]) AND ("ROLL_IO".Input[123, 6] OR "ROLL_State".M[70, 3] OR "ROLL_State".M[70, 5] OR "ROLL_State".M[70, 6]) AND ("ROLL_State".M[74, 0] OR "ROLL_State".M[74, 4]));
    "ROLL_State".M[74, 5] := #r;
    // PB16, STEP 5 network 6
    #r := ((NOT "ROLL_IO".Input[11, 0]) AND (NOT "ROLL_IO".Input[11, 1]) AND (NOT "ROLL_IO".Input[11, 2]) AND (NOT "ROLL_IO".Input[11, 3]) AND (NOT "ROLL_IO".Input[11, 4]) AND (NOT "ROLL_IO".Input[119, 6]) AND (NOT "ROLL_IO".Input[119, 7]) AND (NOT "ROLL_IO".Input[120, 0]) AND (NOT "ROLL_IO".Input[120, 1]));
    "ROLL_State".M[75, 2] := #r;
    // PB16, STEP 5 network 7
    #r := (("ROLL_State".M[190, 6] AND "ROLL_State".M[23, 1] AND "ROLL_State".M[75, 3]) OR "ROLL_State".M[75, 2]);
    "ROLL_State".M[75, 3] := #r;
    // PB16, STEP 5 network 8
    #r := ((((NOT "ROLL_IO".Input[11, 0]) AND (NOT "ROLL_IO".Input[11, 1]) AND (NOT "ROLL_IO".Input[11, 2]) AND (NOT "ROLL_IO".Input[11, 3]) AND (NOT "ROLL_IO".Input[11, 4]) AND (NOT "ROLL_IO".Input[119, 6]) AND (NOT "ROLL_IO".Input[119, 7]) AND (NOT "ROLL_IO".Input[120, 0]) AND (NOT "ROLL_IO".Input[120, 1]) AND "ROLL_IO".Input[13, 3]) OR "ROLL_State".M[63, 1]) AND ((NOT "ROLL_IO".Input[11, 6]) OR (NOT "ROLL_State".M[75, 3]) OR "ROLL_State".M[75, 2]) AND "ROLL_IO".Input[0, 1] AND "ROLL_IO".Input[12, 5] AND "ROLL_State".M[190, 6] AND "ROLL_State".M[23, 1]);
    "ROLL_State".M[75, 4] := #r;
    // PB16, STEP 5 network 9
    #r := ((((NOT "ROLL_IO".Input[11, 0]) AND (NOT "ROLL_IO".Input[11, 1]) AND (NOT "ROLL_IO".Input[11, 2]) AND (NOT "ROLL_IO".Input[11, 3]) AND (NOT "ROLL_IO".Input[11, 4]) AND (NOT "ROLL_IO".Input[119, 6]) AND (NOT "ROLL_IO".Input[119, 7]) AND (NOT "ROLL_IO".Input[120, 0]) AND (NOT "ROLL_IO".Input[120, 1]) AND "ROLL_IO".Input[13, 3]) OR "ROLL_State".M[63, 1]) AND (((NOT "ROLL_State".M[190, 6]) AND "ROLL_State".M[190, 5] AND "ROLL_State".M[23, 1]) OR "ROLL_State".M[74, 0]) AND "ROLL_IO".Input[0, 1]);
    "ROLL_State".M[75, 5] := #r;
    // PB16, STEP 5 network 10
    #r := (((NOT "ROLL_IO".Input[11, 0]) AND (("ROLL_IO".Input[0, 1] AND "ROLL_State".M[190, 5] AND "ROLL_State".M[23, 1]) OR "ROLL_State".M[74, 0]) AND "ROLL_State".M[63, 1]) OR ("ROLL_IO".Input[0, 1] AND "ROLL_State".M[190, 6] AND "ROLL_State".M[23, 1] AND "ROLL_State".M[75, 2]));
    "ROLL_State".M[75, 6] := #r;
    // PB16, STEP 5 network 11
    #r := ((NOT "ROLL_IO".Input[11, 0]) AND "ROLL_IO".Input[11, 6] AND "ROLL_State".M[190, 5] AND "ROLL_State".M[23, 0]);
    "ROLL_State".M[76, 0] := #r;
    // PB16, STEP 5 network 12
    #r := (((NOT "ROLL_IO".Input[11, 0]) AND "ROLL_State".M[74, 0]) OR ("ROLL_IO".Input[11, 0] AND "ROLL_IO".Input[11, 6] AND "ROLL_State".M[190, 6] AND "ROLL_State".M[23, 0]));
    "ROLL_State".M[76, 1] := #r;
    // PB16, STEP 5 network 13
    #r := (("ROLL_State".M[76, 0] OR "ROLL_State".M[76, 1]) AND "ROLL_IO".Input[0, 1]);
    "ROLL_State".M[76, 2] := #r;
    // PB16, STEP 5 network 14
    #r := ((NOT "ROLL_IO".Input[12, 1]) AND (NOT "ROLL_IO".Input[12, 5]));
    "ROLL_State".M[240, 0] := #r;
    // PB16, STEP 5 network 15
    #r := (("ROLL_State".M[190, 6] AND "ROLL_State".M[23, 0] AND "ROLL_State".M[77, 1]) OR "ROLL_State".M[240, 0]);
    "ROLL_State".M[77, 1] := #r;
    // PB16, STEP 5 network 16
    #r := ((((NOT "ROLL_IO".Input[12, 1]) AND ("ROLL_IO".Input[11, 1] OR "ROLL_IO".Input[11, 2] OR "ROLL_IO".Input[11, 3] OR "ROLL_IO".Input[11, 4] OR "ROLL_IO".Input[119, 6] OR "ROLL_IO".Input[119, 7] OR "ROLL_IO".Input[120, 0] OR "ROLL_IO".Input[120, 1])) OR (NOT "ROLL_IO".Input[12, 7])) AND ((NOT "ROLL_IO".Input[12, 7]) OR (NOT "ROLL_State".M[77, 1]) OR "ROLL_State".M[240, 0]) AND "ROLL_IO".Input[0, 1] AND "ROLL_IO".Input[11, 6] AND "ROLL_State".M[190, 6] AND "ROLL_State".M[23, 0]);
    "ROLL_State".M[77, 2] := #r;
    // PB16, STEP 5 network 17
    #r := (((NOT "ROLL_State".M[6, 0]) AND (NOT "ROLL_State".M[6, 2]) AND ("ROLL_IO".Input[11, 1] OR "ROLL_IO".Input[11, 2] OR "ROLL_IO".Input[11, 3] OR "ROLL_IO".Input[11, 4] OR "ROLL_IO".Input[119, 6] OR "ROLL_IO".Input[119, 7] OR "ROLL_IO".Input[120, 0])) OR "ROLL_IO".Input[11, 4]);
    "ROLL_State".M[76, 4] := #r;
    // PB16, STEP 5 network 18
    #r := ((NOT "ROLL_State".M[190, 5]) AND "ROLL_State".M[190, 6] AND "ROLL_State".M[23, 0] AND "ROLL_State".M[76, 4] AND "ROLL_State".M[77, 2]);
    "ROLL_State".M[76, 5] := #r;
    // PB16, STEP 5 network 19
    #r := ((((NOT "ROLL_State".M[190, 6]) AND "ROLL_State".M[190, 5] AND "ROLL_State".M[23, 0]) OR "ROLL_State".M[74, 0]) AND (("ROLL_IO".Input[124, 2] AND "ROLL_IO".Input[124, 5]) OR "ROLL_State".M[0, 4]) AND "ROLL_IO".Input[11, 0] AND "ROLL_State".M[63, 1]);
    "ROLL_State".M[76, 6] := #r;
    // PB16, STEP 5 network 20
    #r := (((((NOT "ROLL_IO".Input[12, 1]) OR (NOT "ROLL_IO".Input[12, 7])) AND "ROLL_State".M[76, 6]) OR "ROLL_State".M[76, 5]) AND "ROLL_IO".Input[0, 1] AND "ROLL_IO".Input[11, 6]);
    "ROLL_State".M[77, 0] := #r;
    // PB16, STEP 5 network 21
    #r := (((NOT "ROLL_IO".Input[11, 0]) AND (NOT "ROLL_IO".Input[12, 5]) AND "ROLL_State".M[190, 5]) OR ((NOT "ROLL_IO".Input[12, 1]) AND "ROLL_IO".Input[11, 0] AND "ROLL_State".M[190, 6]));
    "ROLL_State".M[240, 0] := #r;
    // PB16, STEP 5 network 22
    #r := ((NOT "ROLL_IO".Input[12, 1]) AND ("ROLL_IO".Input[11, 1] OR "ROLL_IO".Input[11, 2] OR "ROLL_IO".Input[11, 3] OR "ROLL_IO".Input[11, 4] OR "ROLL_IO".Input[119, 6] OR "ROLL_IO".Input[119, 7] OR "ROLL_IO".Input[120, 0]));
    "ROLL_State".M[240, 1] := #r;
    // PB16, STEP 5 network 23
    #r := ((NOT "ROLL_IO".Input[12, 1]) AND "ROLL_IO".Input[11, 0]);
    "ROLL_State".M[240, 2] := #r;
    // PB16, STEP 5 network 24
    #r := ((("ROLL_State".M[240, 1] OR "ROLL_State".M[240, 2]) AND "ROLL_State".M[77, 0]) OR ("ROLL_State".M[240, 0] AND "ROLL_State".M[76, 2]));
    "ROLL_State".M[76, 7] := #r;
    // PB16, STEP 5 network 25
    #r := ((NOT "ROLL_IO".Output[113, 3]) AND (NOT "ROLL_State".M[70, 2]) AND (NOT "ROLL_State".M[70, 3]) AND "ROLL_IO".Input[0, 1] AND "ROLL_IO".Input[11, 0] AND "ROLL_IO".Input[12, 1] AND "ROLL_IO".Input[12, 7] AND "ROLL_IO".Input[124, 5]);
    "ROLL_State".M[77, 3] := #r;
    // PB16, STEP 5 network 26
    #r := ((NOT "ROLL_State".M[77, 6]) AND (((NOT "ROLL_State".M[190, 6]) AND "ROLL_State".M[190, 5] AND "ROLL_State".M[22, 0]) OR "ROLL_State".M[74, 0]) AND "ROLL_IO".Output[113, 2] AND "ROLL_State".M[77, 3]);
    "ROLL_State".M[77, 4] := #r;
    // PB16, STEP 5 network 27
    #r := ((NOT "ROLL_State".M[190, 5]) AND (NOT "ROLL_State".M[77, 4]) AND "ROLL_State".M[190, 6] AND "ROLL_State".M[22, 0] AND "ROLL_State".M[77, 3]);
    "ROLL_State".M[77, 6] := #r;
    // PB16, STEP 5 network 28
    #r := ((NOT "ROLL_IO".Input[124, 5]) AND (NOT "ROLL_State".M[70, 3]) AND (((NOT "ROLL_IO".Input[124, 4]) AND "ROLL_State".M[20, 2] AND "ROLL_State".M[74, 0]) OR ((NOT "ROLL_State".M[190, 5]) AND "ROLL_IO".Input[0, 1] AND "ROLL_State".M[190, 6] AND "ROLL_State".M[22, 1])) AND "ROLL_IO".Input[124, 1]);
    "ROLL_State".M[77, 7] := #r;
    // PB16, STEP 5 network 29
    #r := ((NOT "ROLL_IO".Input[124, 4]) AND (NOT "ROLL_State".M[70, 3]) AND (((NOT "ROLL_State".M[15, 1]) AND "ROLL_State".M[20, 1] AND "ROLL_State".M[74, 0]) OR ((NOT "ROLL_State".M[190, 6]) AND "ROLL_IO".Input[0, 1] AND "ROLL_State".M[190, 5] AND "ROLL_State".M[22, 1])) AND "ROLL_IO".Input[124, 1]);
    "ROLL_State".M[78, 0] := #r;
    // PB16, STEP 5 network 30
    #r := ((("ROLL_State".M[22, 3] OR "ROLL_State".M[22, 4]) AND "ROLL_IO".Input[0, 1] AND "ROLL_State".M[190, 6]) OR ("ROLL_IO".Input[123, 5] AND "ROLL_State".M[74, 0]));
    IF #r THEN "ROLL_State".M[78, 4] := TRUE; END_IF;
    #r := (((NOT "ROLL_IO".Output[113, 3]) AND (NOT "ROLL_IO".Input[123, 4]) AND "ROLL_State".M[74, 0]) OR ((NOT "ROLL_IO".Output[113, 3]) AND "ROLL_IO".Input[0, 1] AND "ROLL_State".M[190, 5] AND "ROLL_State".M[22, 3]) OR (NOT "ROLL_IO".Input[0, 1]));
    IF #r THEN "ROLL_State".M[78, 4] := FALSE; END_IF;
    // PB16, STEP 5 network 31
    #r := ((NOT "ROLL_IO".Input[123, 5]) AND (NOT "ROLL_IO".Input[123, 6]) AND (NOT "ROLL_State".M[16, 0]) AND (NOT "ROLL_State".M[16, 4]) AND (NOT "ROLL_State".M[9, 1]) AND ((NOT "ROLL_IO".Input[123, 4]) OR "ROLL_State".M[190, 1]));
    "ROLL_State".M[78, 5] := #r;
    // PB16, STEP 5 network 32
    #r := (((NOT "ROLL_IO".Input[124, 2]) AND (NOT "ROLL_State".M[190, 5]) AND (NOT "ROLL_State".M[70, 3]) AND "ROLL_IO".Input[0, 1] AND "ROLL_IO".Input[124, 1] AND "ROLL_IO".Input[124, 4] AND "ROLL_State".M[190, 6] AND "ROLL_State".M[22, 4]) OR ("ROLL_State".M[70, 2] AND "ROLL_State".M[74, 0]));
    IF #r THEN "ROLL_State".M[78, 6] := TRUE; END_IF;
    #r := (((NOT "ROLL_State".M[70, 2]) AND ((NOT "ROLL_IO".Input[124, 1]) OR (NOT "ROLL_IO".Input[124, 4])) AND "ROLL_State".M[20, 2] AND "ROLL_State".M[74, 0]) OR ((NOT "ROLL_State".M[70, 2]) AND "ROLL_IO".Input[0, 1] AND "ROLL_State".M[190, 5] AND "ROLL_State".M[22, 4]) OR ((NOT "ROLL_State".M[70, 2]) AND "ROLL_State".M[20, 1] AND "ROLL_State".M[74, 0]) OR (NOT "ROLL_IO".Input[0, 1]) OR "ROLL_State".M[70, 0]);
    IF #r THEN "ROLL_State".M[78, 6] := FALSE; END_IF;
    // PB16, STEP 5 network 33
    #r := (((NOT "ROLL_State".M[70, 2]) AND (("ROLL_IO".Input[124, 5] AND "ROLL_State".M[20, 2]) OR "ROLL_State".M[20, 1]) AND "ROLL_State".M[74, 0]) OR ((NOT "ROLL_State".M[70, 2]) AND "ROLL_IO".Input[0, 1] AND "ROLL_State".M[190, 5] AND "ROLL_State".M[22, 4]));
    IF #r THEN "ROLL_State".M[78, 7] := TRUE; END_IF;
    #r := ((NOT "ROLL_IO".Input[0, 1]) OR "ROLL_State".M[70, 0] OR "ROLL_State".M[78, 6]);
    IF #r THEN "ROLL_State".M[78, 7] := FALSE; END_IF;
    // PB16, STEP 5 network 34
    RETURN;
END_FUNCTION

FUNCTION "ROLL_PB17" : Void
{ S7_Optimized_Access := 'TRUE' }
VERSION : 0.1
VAR_TEMP
    r : Bool;
    a1 : Word;
    a2 : Word;
    activeDataBlock : Int;
    comparisonResults : Array[0..0] of Bool;
END_VAR
BEGIN
    #r := FALSE;
    #a1 := W#16#0000;
    #a2 := W#16#0000;
    #activeDataBlock := 0;
    // PB17, STEP 5 network 1
    #r := ((NOT "ROLL_State".M[70, 1]) AND "ROLL_State".M[3, 3]);
    "ROLL_State".M[70, 0] := #r;
    // PB17, STEP 5 network 2
    #r := "ROLL_State".M[70, 0];
    IF #r THEN "ROLL_State".M[70, 1] := TRUE; END_IF;
    #r := "ROLL_IO".Input[0, 2];
    IF #r THEN "ROLL_State".M[70, 1] := FALSE; END_IF;
    // PB17, STEP 5 network 3
    #r := ((("ROLL_IO".Input[0, 1] AND "ROLL_State".M[74, 1]) OR ("ROLL_IO".Input[0, 2] AND "ROLL_State".M[64, 0])) AND "ROLL_State".M[29, 1]);
    "ROLL_IO".Output[112, 0] := #r;
    // PB17, STEP 5 network 4
    #r := ((("ROLL_IO".Input[0, 1] AND "ROLL_State".M[74, 5]) OR ("ROLL_IO".Input[0, 2] AND "ROLL_State".M[64, 1])) AND "ROLL_State".M[29, 1]);
    "ROLL_IO".Output[112, 5] := #r;
    // PB17, STEP 5 network 5
    #r := (((("ROLL_IO".Input[0, 1] AND "ROLL_State".M[78, 4]) OR ("ROLL_IO".Input[0, 2] AND "ROLL_State".M[64, 4])) AND "ROLL_State".M[29, 0]) OR ("ROLL_IO".Output[113, 1] AND "ROLL_IO".Output[113, 3]));
    "ROLL_IO".Output[113, 1] := #r;
    // PB17, STEP 5 network 6
    #r := (((NOT "ROLL_State".M[71, 4]) AND "ROLL_State".M[71, 3]) OR ((("ROLL_IO".Input[0, 1] AND "ROLL_State".M[78, 6]) OR ("ROLL_IO".Input[0, 2] AND "ROLL_State".M[64, 5])) AND "ROLL_State".M[29, 0]));
    "ROLL_State".M[71, 3] := #r;
    // PB17, STEP 5 network 7
    #r := "ROLL_State".M[71, 3];
    "ROLL_IO".Output[113, 3] := #r;
    // PB17, STEP 5 network 8
    #r := (((NOT "ROLL_State".M[71, 3]) AND "ROLL_State".M[71, 4]) OR ((((NOT "ROLL_State".M[64, 5]) AND ((NOT "ROLL_State".M[20, 2]) OR "ROLL_IO".Input[124, 5]) AND "ROLL_IO".Input[0, 2]) OR ("ROLL_IO".Input[0, 1] AND "ROLL_State".M[78, 7])) AND "ROLL_State".M[29, 0]));
    "ROLL_State".M[71, 4] := #r;
    // PB17, STEP 5 network 9
    #r := "ROLL_State".M[71, 4];
    "ROLL_IO".Output[113, 2] := #r;
    // PB17, STEP 5 network 10
    #r := (("ROLL_IO".Input[0, 1] AND "ROLL_State".M[75, 4]) OR ("ROLL_IO".Input[0, 2] AND "ROLL_State".M[35, 2] AND "ROLL_State".M[65, 0]));
    "ROLL_State".M[79, 5] := #r;
    // PB17, STEP 5 network 11
    #r := ((NOT "ROLL_IO".Output[23, 0]) AND (NOT "ROLL_IO".Output[23, 4]) AND (NOT "ROLL_State".M[10, 3]) AND (NOT "ROLL_State".M[5, 0]) AND ((NOT "ROLL_IO".Input[11, 4]) OR (NOT "ROLL_IO".Input[11, 6])) AND "ROLL_IO".Input[11, 7] AND "ROLL_IO".Input[12, 5] AND "ROLL_IO".Input[12, 7] AND "ROLL_IO".Input[14, 0] AND "ROLL_State".M[29, 0] AND "ROLL_State".M[79, 5]);
    "ROLL_IO".Output[23, 1] := #r;
    // PB17, STEP 5 network 12
    #r := (("ROLL_IO".Input[0, 1] AND "ROLL_State".M[75, 5]) OR ("ROLL_IO".Input[0, 2] AND "ROLL_State".M[35, 2] AND "ROLL_State".M[65, 5]));
    "ROLL_State".M[79, 6] := #r;
    // PB17, STEP 5 network 13
    #r := ((NOT "ROLL_IO".Output[23, 1]) AND (NOT "ROLL_IO".Output[23, 4]) AND (NOT "ROLL_State".M[10, 2]) AND (NOT "ROLL_State".M[5, 0]) AND (((NOT "ROLL_IO".Input[119, 0]) AND "ROLL_State".M[0, 3]) OR (NOT "ROLL_IO".Input[11, 0]) OR (NOT "ROLL_IO".Input[11, 6])) AND "ROLL_IO".Input[11, 7] AND "ROLL_IO".Input[12, 5] AND "ROLL_IO".Input[12, 7] AND "ROLL_IO".Input[14, 0] AND "ROLL_State".M[29, 0] AND "ROLL_State".M[79, 6]);
    "ROLL_IO".Output[23, 0] := #r;
    // PB17, STEP 5 network 14
    #r := ((("ROLL_IO".Input[0, 1] AND "ROLL_State".M[75, 6]) OR ("ROLL_IO".Input[0, 2] AND "ROLL_State".M[35, 2] AND "ROLL_State".M[65, 6])) AND ("ROLL_IO".Output[23, 0] OR "ROLL_IO".Output[23, 1]));
    "ROLL_IO".Output[23, 3] := #r;
    // PB17, STEP 5 network 15
    #r := ((NOT "ROLL_IO".Output[23, 3]) AND ("ROLL_IO".Output[23, 0] OR "ROLL_IO".Output[23, 1]) AND ("ROLL_IO".Input[0, 1] OR "ROLL_State".M[31, 5]) AND "ROLL_State".M[29, 0]);
    "ROLL_IO".Output[23, 2] := #r;
    // PB17, STEP 5 network 16
    #r := (("ROLL_IO".Input[0, 1] AND "ROLL_State".M[76, 2]) OR ("ROLL_IO".Input[0, 2] AND "ROLL_State".M[35, 2] AND "ROLL_State".M[66, 4]));
    "ROLL_State".M[80, 0] := #r;
    // PB17, STEP 5 network 17
    #r := ((NOT "ROLL_IO".Output[23, 4]) AND (NOT "ROLL_State".M[10, 1]) AND (NOT "ROLL_State".M[5, 2]) AND (NOT "ROLL_State".M[9, 0]) AND ((NOT "ROLL_IO".Input[12, 5]) OR (NOT "ROLL_IO".Input[12, 7])) AND ("ROLL_IO".Input[124, 2] OR "ROLL_State".M[0, 4]) AND "ROLL_IO".Input[13, 0] AND "ROLL_IO".Input[13, 7] AND "ROLL_IO".Input[14, 0] AND "ROLL_State".M[29, 0] AND "ROLL_State".M[80, 0]);
    "ROLL_IO".Output[23, 5] := #r;
    // PB17, STEP 5 network 18
    #r := (("ROLL_IO".Input[0, 1] AND "ROLL_State".M[77, 0]) OR ("ROLL_IO".Input[0, 2] AND "ROLL_State".M[35, 2] AND "ROLL_State".M[66, 7]));
    "ROLL_State".M[80, 1] := #r;
    // PB17, STEP 5 network 19
    #r := "ROLL_IO".Input[12, 5];
    IF #r THEN "ROLL_State".M[80, 2] := TRUE; END_IF;
    #r := "ROLL_IO".Input[12, 1];
    IF #r THEN "ROLL_State".M[80, 2] := FALSE; END_IF;
    // PB17, STEP 5 network 20
    #r := (((("ROLL_IO".Input[11, 1] OR "ROLL_IO".Input[11, 2] OR "ROLL_IO".Input[11, 3] OR "ROLL_IO".Input[11, 4] OR "ROLL_IO".Input[119, 6] OR "ROLL_IO".Input[119, 7] OR "ROLL_IO".Input[120, 0] OR "ROLL_IO".Input[120, 1]) AND "ROLL_IO".Input[12, 1]) OR ("ROLL_IO".Input[11, 0] AND "ROLL_IO".Input[12, 1])) AND "ROLL_IO".Input[12, 7]);
    "ROLL_State".M[80, 6] := #r;
    // PB17, STEP 5 network 21
    #r := (("ROLL_IO".Input[11, 0] OR "ROLL_IO".Input[11, 1] OR "ROLL_IO".Input[11, 2] OR "ROLL_IO".Input[11, 3] OR "ROLL_IO".Input[11, 4] OR "ROLL_IO".Input[119, 6] OR "ROLL_IO".Input[119, 7] OR "ROLL_IO".Input[120, 0] OR "ROLL_IO".Input[120, 1]) AND "ROLL_IO".Input[12, 5] AND "ROLL_IO".Input[12, 7]);
    "ROLL_State".M[80, 7] := #r;
    // PB17, STEP 5 network 22
    #r := ((NOT "ROLL_IO".Output[23, 0]) AND (NOT "ROLL_IO".Output[23, 1]) AND (NOT "ROLL_IO".Output[23, 5]) AND (NOT "ROLL_State".M[10, 0]) AND (NOT "ROLL_State".M[5, 2]) AND (NOT "ROLL_State".M[80, 6]) AND ("ROLL_IO".Input[124, 2] OR "ROLL_State".M[0, 4]) AND "ROLL_IO".Input[13, 0] AND "ROLL_IO".Input[14, 0] AND "ROLL_State".M[29, 0] AND "ROLL_State".M[80, 1]);
    "ROLL_IO".Output[23, 4] := #r;
    // PB17, STEP 5 network 23
    #r := ((NOT "ROLL_State".M[68, 2]) AND (((NOT "ROLL_IO".Input[12, 5]) AND "ROLL_IO".Output[23, 5]) OR ("ROLL_IO".Output[23, 4] AND "ROLL_State".M[80, 2])));
    "ROLL_IO".Output[23, 7] := #r;
    // PB17, STEP 5 network 24
    #r := ((NOT "ROLL_IO".Output[23, 7]) AND ("ROLL_IO".Output[23, 4] OR "ROLL_IO".Output[23, 5]));
    "ROLL_IO".Output[23, 6] := #r;
    // PB17, STEP 5 network 25
    #r := (("ROLL_IO".Input[0, 1] AND "ROLL_State".M[77, 6]) OR ("ROLL_IO".Input[0, 2] AND "ROLL_State".M[35, 2] AND "ROLL_State".M[67, 0]));
    "ROLL_State".M[80, 3] := #r;
    // PB17, STEP 5 network 26
    #r := ((NOT "ROLL_IO".Output[112, 1]) AND (NOT "ROLL_IO".Output[113, 3]) AND (NOT "ROLL_IO".Input[124, 2]) AND (NOT "ROLL_State".M[10, 5]) AND (NOT "ROLL_State".M[70, 2]) AND (NOT "ROLL_State".M[9, 3]) AND "ROLL_IO".Input[11, 0] AND "ROLL_IO".Input[11, 6] AND "ROLL_IO".Input[12, 1] AND "ROLL_IO".Input[12, 7] AND "ROLL_State".M[29, 0] AND "ROLL_State".M[80, 3]);
    "ROLL_IO".Output[112, 2] := #r;
    // PB17, STEP 5 network 27
    #r := (("ROLL_IO".Input[0, 1] AND "ROLL_State".M[77, 4]) OR ("ROLL_IO".Input[0, 2] AND "ROLL_State".M[35, 2] AND "ROLL_State".M[67, 1]));
    "ROLL_State".M[80, 4] := #r;
    // PB17, STEP 5 network 28
    #r := ((NOT "ROLL_IO".Output[112, 2]) AND (NOT "ROLL_IO".Output[113, 3]) AND (NOT "ROLL_IO".Input[124, 1]) AND (NOT "ROLL_State".M[10, 4]) AND (NOT "ROLL_State".M[70, 2]) AND (NOT "ROLL_State".M[70, 3]) AND (NOT "ROLL_State".M[9, 3]) AND "ROLL_IO".Input[11, 0] AND "ROLL_IO".Input[11, 6] AND "ROLL_IO".Input[12, 1] AND "ROLL_IO".Input[12, 7] AND "ROLL_State".M[29, 0] AND "ROLL_State".M[80, 4]);
    "ROLL_IO".Output[112, 1] := #r;
    // PB17, STEP 5 network 29
    #r := ((("ROLL_IO".Input[0, 1] AND "ROLL_State".M[77, 7]) OR ("ROLL_IO".Input[0, 2] AND "ROLL_State".M[35, 2] AND "ROLL_State".M[67, 5])) AND "ROLL_State".M[29, 0]);
    "ROLL_IO".Output[112, 4] := #r;
    // PB17, STEP 5 network 30
    #r := ((("ROLL_IO".Input[0, 1] AND "ROLL_State".M[78, 0]) OR ("ROLL_IO".Input[0, 2] AND "ROLL_State".M[35, 2] AND "ROLL_State".M[67, 6])) AND "ROLL_State".M[29, 0]);
    "ROLL_IO".Output[112, 3] := #r;
    // PB17, STEP 5 network 31
    #r := ((NOT "ROLL_State".M[16, 0]) AND (NOT "ROLL_State".M[16, 1]) AND (NOT "ROLL_State".M[16, 2]) AND (NOT "ROLL_State".M[16, 4]) AND "ROLL_State".M[37, 2]);
    "ROLL_State".M[81, 4] := #r;
    // PB17, STEP 5 network 32
    RETURN;
END_FUNCTION

FUNCTION "ROLL_PB18" : Void
{ S7_Optimized_Access := 'TRUE' }
VERSION : 0.1
VAR_TEMP
    r : Bool;
    a1 : Word;
    a2 : Word;
    activeDataBlock : Int;
    comparisonResults : Array[0..0] of Bool;
END_VAR
BEGIN
    #r := FALSE;
    #a1 := W#16#0000;
    #a2 := W#16#0000;
    #activeDataBlock := 0;
    // PB18, STEP 5 network 1
    #r := ("ROLL_State".M[70, 2] OR "ROLL_State".M[70, 3] OR "ROLL_State".M[70, 4] OR "ROLL_State".M[70, 6] OR "ROLL_State".M[71, 0]);
    "ROLL_State".M[80, 5] := #r;
    // PB18, STEP 5 network 2
    #r := (((NOT "ROLL_IO".Output[112, 0]) AND (NOT "ROLL_IO".Output[112, 5]) AND "ROLL_State".M[20, 5]) OR ((NOT "ROLL_IO".Output[112, 0]) AND "ROLL_State".M[20, 3]) OR ((NOT "ROLL_IO".Output[112, 5]) AND "ROLL_State".M[20, 4]) OR ((NOT "ROLL_IO".Output[17, 7]) AND "ROLL_State".M[20, 7]) OR (("ROLL_State".M[20, 1] OR "ROLL_State".M[20, 2]) AND "ROLL_State".M[28, 4]));
    "ROLL_State".M[250, 0] := #r;
    // PB18, STEP 5 network 3
    #r := (((NOT "ROLL_IO".Output[113, 0]) AND "ROLL_State".M[22, 2]) OR ((NOT "ROLL_IO".Output[113, 1]) AND "ROLL_State".M[22, 3]) OR ((NOT "ROLL_IO".Output[113, 3]) AND "ROLL_IO".Output[113, 2] AND "ROLL_State".M[22, 4]) OR ((NOT "ROLL_IO".Output[113, 5]) AND "ROLL_IO".Output[113, 4] AND "ROLL_State".M[22, 5]) OR ("ROLL_IO".Input[124, 1] AND "ROLL_State".M[22, 0]) OR ("ROLL_IO".Input[124, 4] AND "ROLL_State".M[22, 1]) OR "ROLL_State".M[250, 0]);
    "ROLL_State".M[250, 0] := #r;
    // PB18, STEP 5 network 4
    #r := ((("ROLL_IO".Input[11, 1] OR "ROLL_IO".Input[11, 2] OR "ROLL_IO".Input[11, 3] OR "ROLL_IO".Input[11, 4] OR "ROLL_IO".Input[119, 6] OR "ROLL_IO".Input[119, 7] OR "ROLL_IO".Input[120, 0] OR "ROLL_IO".Input[120, 1]) AND "ROLL_IO".Input[12, 5] AND "ROLL_IO".Input[12, 7] AND "ROLL_State".M[23, 0]) OR (("ROLL_State".M[23, 2] OR "ROLL_State".M[23, 3]) AND "ROLL_State".M[63, 1]) OR ("ROLL_IO".Input[11, 0] AND "ROLL_IO".Input[11, 6] AND "ROLL_State".M[23, 1]) OR ("ROLL_IO".Input[11, 0] AND "ROLL_IO".Input[12, 1] AND "ROLL_IO".Input[12, 7] AND "ROLL_State".M[23, 0]) OR "ROLL_State".M[250, 0]);
    "ROLL_State".M[250, 0] := #r;
    // PB18, STEP 5 network 5
    #r := (((NOT "ROLL_IO".Output[20, 1]) AND "ROLL_State".M[24, 1]) OR "ROLL_State".M[250, 0]);
    "ROLL_State".M[250, 0] := #r;
    // PB18, STEP 5 network 6
    #r := ((((NOT "ROLL_IO".Output[20, 4]) OR (NOT "ROLL_IO".Output[22, 6])) AND "ROLL_State".M[25, 0]) OR "ROLL_State".M[250, 0]);
    "ROLL_State".M[250, 0] := #r;
    // PB18, STEP 5 network 7
    #r := (((NOT "ROLL_IO".Output[20, 5]) AND "ROLL_State".M[26, 6]) OR ((NOT "ROLL_IO".Output[20, 6]) AND "ROLL_State".M[26, 0]) OR ((NOT "ROLL_IO".Output[21, 4]) AND "ROLL_State".M[26, 5]) OR "ROLL_State".M[250, 0]);
    "ROLL_State".M[250, 0] := #r;
    // PB18, STEP 5 network 8
    #r := (((NOT "ROLL_IO".Output[20, 6]) AND "ROLL_State".M[27, 4]) OR ((NOT "ROLL_IO".Output[21, 6]) AND "ROLL_State".M[27, 5]) OR ((NOT "ROLL_State".M[80, 5]) AND "ROLL_State".M[27, 7]) OR "ROLL_State".M[250, 0]);
    "ROLL_State".M[250, 0] := #r;
    // PB18, STEP 5 network 9
    #r := ((("ROLL_IO".Output[112, 0] OR "ROLL_IO".Output[112, 5]) AND "ROLL_State".M[20, 5]) OR ("ROLL_IO".Output[112, 0] AND "ROLL_State".M[20, 3]) OR ("ROLL_IO".Output[112, 5] AND "ROLL_State".M[20, 4]) OR ("ROLL_IO".Output[17, 7] AND "ROLL_State".M[20, 7]));
    "ROLL_State".M[252, 0] := #r;
    // PB18, STEP 5 network 10
    #r := (((NOT "ROLL_IO".Output[113, 2]) AND "ROLL_IO".Output[113, 3] AND "ROLL_State".M[22, 4]) OR ((NOT "ROLL_IO".Output[113, 4]) AND "ROLL_IO".Output[113, 5] AND "ROLL_State".M[22, 5]) OR ("ROLL_IO".Output[113, 0] AND "ROLL_State".M[22, 2]) OR ("ROLL_IO".Output[113, 1] AND "ROLL_State".M[22, 3]) OR ("ROLL_IO".Input[124, 2] AND "ROLL_State".M[22, 0]) OR ("ROLL_IO".Input[124, 5] AND "ROLL_State".M[22, 1]) OR "ROLL_State".M[252, 0]);
    "ROLL_State".M[252, 0] := #r;
    // PB18, STEP 5 network 11
    #r := (((NOT "ROLL_IO".Output[23, 1]) AND ("ROLL_IO".Input[11, 1] OR "ROLL_IO".Input[11, 2] OR "ROLL_IO".Input[11, 3] OR "ROLL_IO".Input[11, 4] OR "ROLL_IO".Input[119, 6] OR "ROLL_IO".Input[119, 7] OR "ROLL_IO".Input[120, 0] OR "ROLL_IO".Input[120, 1]) AND "ROLL_IO".Input[11, 6] AND "ROLL_State".M[23, 1]) OR ((NOT "ROLL_State".M[63, 1]) AND ("ROLL_State".M[23, 2] OR "ROLL_State".M[23, 3])) OR (((("ROLL_IO".Input[11, 1] OR "ROLL_IO".Input[11, 2] OR "ROLL_IO".Input[11, 3] OR "ROLL_IO".Input[11, 4] OR "ROLL_IO".Input[119, 6] OR "ROLL_IO".Input[119, 7] OR "ROLL_IO".Input[120, 0] OR "ROLL_IO".Input[120, 1]) AND "ROLL_IO".Input[12, 1]) OR ("ROLL_IO".Input[11, 0] AND "ROLL_IO".Input[12, 5])) AND "ROLL_IO".Input[12, 7] AND "ROLL_State".M[23, 0]) OR "ROLL_State".M[252, 0]);
    "ROLL_State".M[252, 0] := #r;
    // PB18, STEP 5 network 12
    #r := (("ROLL_IO".Output[20, 1] AND "ROLL_State".M[24, 1]) OR "ROLL_State".M[252, 0]);
    "ROLL_State".M[252, 0] := #r;
    // PB18, STEP 5 network 13
    #r := (("ROLL_IO".Output[20, 4] AND "ROLL_IO".Output[22, 6] AND "ROLL_State".M[25, 0]) OR "ROLL_State".M[252, 0]);
    "ROLL_State".M[252, 0] := #r;
    // PB18, STEP 5 network 14
    #r := (("ROLL_IO".Output[20, 6] AND "ROLL_State".M[26, 0]) OR "ROLL_State".M[252, 0]);
    "ROLL_State".M[252, 0] := #r;
    // PB18, STEP 5 network 15
    #r := (("ROLL_IO".Output[20, 5] AND "ROLL_State".M[26, 6]) OR ("ROLL_IO".Output[20, 6] AND "ROLL_State".M[27, 4]) OR ("ROLL_IO".Output[21, 4] AND "ROLL_State".M[26, 5]) OR ("ROLL_IO".Output[21, 6] AND "ROLL_State".M[27, 5]) OR ("ROLL_State".M[27, 7] AND "ROLL_State".M[80, 5]) OR "ROLL_State".M[252, 0]);
    "ROLL_State".M[252, 0] := #r;
    // PB18, STEP 5 network 16
    RETURN;
END_FUNCTION

FUNCTION "ROLL_PB19" : Void
{ S7_Optimized_Access := 'TRUE' }
VERSION : 0.1
VAR_TEMP
    r : Bool;
    a1 : Word;
    a2 : Word;
    activeDataBlock : Int;
    comparisonResults : Array[0..0] of Bool;
END_VAR
BEGIN
    #r := FALSE;
    #a1 := W#16#0000;
    #a2 := W#16#0000;
    #activeDataBlock := 0;
    // PB19, STEP 5 network 1
    #r := ((NOT "ROLL_IO".Input[3, 6]) AND (NOT "ROLL_State".M[5, 6]) AND (NOT "ROLL_State".M[6, 0]) AND (NOT "ROLL_State".M[6, 2]) AND ("ROLL_IO".Input[3, 1] OR "ROLL_State".M[31, 5]) AND "ROLL_IO".Input[5, 2] AND "ROLL_IO".Input[5, 4] AND "ROLL_State".M[4, 1]);
    "ROLL_State".M[82, 0] := #r;
    // PB19, STEP 5 network 2
    #r := ((NOT "ROLL_IO".Input[3, 6]) AND (NOT "ROLL_State".M[12, 0]) AND (NOT "ROLL_State".M[5, 3]) AND (NOT "ROLL_State".M[5, 6]) AND ("ROLL_IO".Input[3, 1] OR "ROLL_State".M[31, 5]) AND "ROLL_IO".Input[8, 3] AND "ROLL_IO".Input[8, 5] AND "ROLL_State".M[4, 1]);
    "ROLL_State".M[82, 2] := #r;
    // PB19, STEP 5 network 3
    #r := ("ROLL_State".M[31, 5] AND "ROLL_State".M[40, 0]);
    IF #r THEN "ROLL_State".M[82, 3] := TRUE; END_IF;
    #r := (NOT "ROLL_State".M[31, 5]);
    IF #r THEN "ROLL_State".M[82, 3] := FALSE; END_IF;
    // PB19, STEP 5 network 4
    #r := ((NOT "ROLL_State".M[110, 1]) AND (NOT "ROLL_State".M[110, 2]) AND "ROLL_State".M[110, 0] AND "ROLL_State".M[110, 3] AND "ROLL_State".M[40, 0]);
    "ROLL_State".M[240, 0] := #r;
    // PB19, STEP 5 network 5
    #r := (((NOT "ROLL_State".M[110, 2]) AND "ROLL_State".M[110, 0] AND "ROLL_State".M[110, 1] AND "ROLL_State".M[110, 3] AND "ROLL_State".M[41, 1]) OR "ROLL_State".M[240, 0]);
    "ROLL_State".M[240, 0] := #r;
    // PB19, STEP 5 network 6
    #r := (((NOT "ROLL_State".M[110, 1]) AND "ROLL_State".M[110, 0] AND "ROLL_State".M[110, 2] AND "ROLL_State".M[110, 3] AND "ROLL_State".M[41, 1]) OR "ROLL_State".M[240, 0]);
    "ROLL_State".M[240, 0] := #r;
    // PB19, STEP 5 network 7
    #r := (("ROLL_State".M[110, 0] AND "ROLL_State".M[110, 1] AND "ROLL_State".M[110, 2] AND "ROLL_State".M[110, 3] AND "ROLL_State".M[41, 1]) OR "ROLL_State".M[240, 0]);
    "ROLL_State".M[240, 0] := #r;
    // PB19, STEP 5 network 8
    #r := ("ROLL_State".M[240, 0] AND "ROLL_State".M[31, 5]);
    IF #r THEN "ROLL_State".M[82, 4] := TRUE; END_IF;
    #r := ((NOT "ROLL_State".M[31, 5]) OR "ROLL_State".M[45, 5]);
    IF #r THEN "ROLL_State".M[82, 4] := FALSE; END_IF;
    // PB19, STEP 5 network 9
    #r := ((NOT "ROLL_IO".Output[17, 3]) AND (NOT "ROLL_State".M[82, 4]) AND (NOT "ROLL_State".S5Timers[91].Q) AND ("ROLL_State".M[82, 3] OR "ROLL_State".S5Timers[22].Q) AND "ROLL_IO".Input[8, 5]);
    "ROLL_IO".Output[17, 2] := #r;
    // PB19, STEP 5 network 10
    #r := ((NOT "ROLL_IO".Output[17, 2]) AND (NOT "ROLL_State".S5Timers[90].Q) AND "ROLL_IO".Input[3, 0] AND "ROLL_IO".Input[8, 5] AND "ROLL_State".M[82, 4]);
    "ROLL_IO".Output[17, 3] := #r;
    // PB19, STEP 5 network 11
    #a2 := #a1;
    #a1 := W#16#3060;
    #r := "ROLL_IO".Output[18, 0];
    "ROLL_TimerOp"(Number := 22, Operation := 1, Signal := #r, Preset := #a1);
    // PB19, STEP 5 network 12
    #a2 := #a1;
    #a1 := W#16#1005;
    #r := "ROLL_IO".Output[17, 2];
    "ROLL_TimerOp"(Number := 90, Operation := 1, Signal := #r, Preset := #a1);
    // PB19, STEP 5 network 13
    #a2 := #a1;
    #a1 := W#16#1040;
    #r := "ROLL_IO".Output[17, 3];
    "ROLL_TimerOp"(Number := 91, Operation := 1, Signal := #r, Preset := #a1);
    // PB19, STEP 5 network 14
    #r := ((NOT "ROLL_State".M[12, 0]) AND (NOT "ROLL_State".M[19, 7]) AND ("ROLL_IO".Output[17, 2] OR "ROLL_IO".Output[17, 3] OR "ROLL_State".S5Timers[90].Q OR "ROLL_State".S5Timers[91].Q) AND ("ROLL_State".M[82, 3] OR "ROLL_State".M[82, 4]) AND "ROLL_IO".Input[8, 3] AND "ROLL_IO".Input[8, 4] AND "ROLL_State".M[82, 2]);
    "ROLL_IO".Output[18, 0] := #r;
    // PB19, STEP 5 network 15
    #r := "ROLL_IO".Output[18, 0];
    "ROLL_IO".Output[18, 1] := #r;
    // PB19, STEP 5 network 16
    #r := ("ROLL_IO".Output[18, 0] AND "ROLL_State".M[82, 4]);
    "ROLL_IO".Output[18, 2] := #r;
    // PB19, STEP 5 network 17
    #r := ("ROLL_IO".Output[18, 0] AND "ROLL_State".M[82, 4]);
    "ROLL_IO".Output[18, 3] := #r;
    // PB19, STEP 5 network 18
    RETURN;
END_FUNCTION

FUNCTION "ROLL_PB20" : Void
{ S7_Optimized_Access := 'TRUE' }
VERSION : 0.1
VAR_TEMP
    r : Bool;
    a1 : Word;
    a2 : Word;
    activeDataBlock : Int;
    comparisonResults : Array[0..0] of Bool;
END_VAR
BEGIN
    #r := FALSE;
    #a1 := W#16#0000;
    #a2 := W#16#0000;
    #activeDataBlock := 0;
    // PB20, STEP 5 network 1
    #activeDataBlock := 15;
    // PB20, STEP 5 network 2
    #r := ((NOT "ROLL_IO".Input[7, 0]) AND (("ROLL_IO".Input[0, 1] AND "ROLL_State".M[190, 6] AND "ROLL_State".M[26, 5] AND "ROLL_State".M[4, 1]) OR ("ROLL_IO".Input[0, 2] AND "ROLL_State".M[0, 3])) AND "ROLL_State".M[4, 1]);
    "ROLL_State".M[8, 0] := #r;
    // PB20, STEP 5 network 3
    #r := ((NOT "ROLL_IO".Input[7, 1]) AND "ROLL_IO".Input[0, 2] AND "ROLL_IO".Input[1, 6] AND "ROLL_State".M[4, 1] AND "ROLL_State".S5Timers[61].Q);
    IF #r THEN "ROLL_State".M[8, 1] := TRUE; END_IF;
    #r := "ROLL_State".M[3, 1];
    IF #r THEN "ROLL_State".M[8, 1] := FALSE; END_IF;
    // PB20, STEP 5 network 4
    #a2 := #a1;
    #a1 := "ROLL_GetDW"(DbNumber := #activeDataBlock, Index := 61);
    #r := ((NOT "ROLL_IO".Input[7, 1]) AND "ROLL_IO".Input[0, 2] AND "ROLL_IO".Input[3, 1]);
    "ROLL_TimerOp"(Number := 61, Operation := 0, Signal := #r, Preset := #a1);
    #r := ("ROLL_State".M[3, 1] AND "ROLL_State".M[4, 1]);
    "ROLL_TimerOp"(Number := 61, Operation := 2, Signal := #r, Preset := #a1);
    // PB20, STEP 5 network 5
    #r := ((NOT "ROLL_IO".Input[7, 2]) AND "ROLL_State".S5Timers[55].Q);
    IF #r THEN "ROLL_State".M[8, 2] := TRUE; END_IF;
    #r := "ROLL_State".M[3, 1];
    IF #r THEN "ROLL_State".M[8, 2] := FALSE; END_IF;
    // PB20, STEP 5 network 6
    #a2 := #a1;
    #a1 := "ROLL_GetDW"(DbNumber := #activeDataBlock, Index := 55);
    #r := ((NOT "ROLL_IO".Input[7, 2]) AND (NOT "ROLL_State".M[8, 2]) AND "ROLL_State".M[4, 1]);
    "ROLL_TimerOp"(Number := 55, Operation := 0, Signal := #r, Preset := #a1);
    // PB20, STEP 5 network 7
    #r := ((NOT "ROLL_IO".Input[7, 3]) AND "ROLL_IO".Output[21, 6] AND "ROLL_State".S5Timers[60].Q);
    IF #r THEN "ROLL_State".M[8, 3] := TRUE; END_IF;
    #r := "ROLL_State".M[3, 1];
    IF #r THEN "ROLL_State".M[8, 3] := FALSE; END_IF;
    // PB20, STEP 5 network 8
    #a2 := #a1;
    #a1 := "ROLL_GetDW"(DbNumber := #activeDataBlock, Index := 60);
    #r := ((NOT "ROLL_IO".Input[7, 3]) AND "ROLL_IO".Output[21, 6] AND "ROLL_IO".Input[3, 1]);
    "ROLL_TimerOp"(Number := 60, Operation := 0, Signal := #r, Preset := #a1);
    // PB20, STEP 5 network 9
    #a2 := #a1;
    #a1 := W#16#2010;
    #r := (NOT "ROLL_IO".Input[7, 4]);
    "ROLL_TimerOp"(Number := 88, Operation := 0, Signal := #r, Preset := #a1);
    // PB20, STEP 5 network 10
    #r := ((NOT "ROLL_IO".Input[7, 4]) AND "ROLL_State".M[4, 1] AND "ROLL_State".S5Timers[88].Q);
    "ROLL_State".M[8, 4] := #r;
    // PB20, STEP 5 network 11
    #r := (("ROLL_State".M[25, 0] OR "ROLL_State".M[25, 1]) AND "ROLL_IO".Input[0, 1] AND "ROLL_State".M[190, 6] AND "ROLL_State".M[4, 1] AND "ROLL_State".S5Timers[96].Q);
    IF #r THEN "ROLL_State".M[8, 5] := TRUE; END_IF;
    #r := "ROLL_State".M[3, 1];
    IF #r THEN "ROLL_State".M[8, 5] := FALSE; END_IF;
    // PB20, STEP 5 network 12
    #r := ((NOT "ROLL_IO".Input[9, 0]) AND ("ROLL_IO".Input[1, 6] OR "ROLL_IO".Input[1, 7]) AND "ROLL_IO".Input[9, 6]);
    IF #r THEN "ROLL_State".M[12, 4] := TRUE; END_IF;
    #r := "ROLL_State".M[3, 1];
    IF #r THEN "ROLL_State".M[12, 4] := FALSE; END_IF;
    // PB20, STEP 5 network 13
    #r := ((NOT "ROLL_IO".Input[9, 3]) AND ("ROLL_IO".Input[1, 6] OR "ROLL_IO".Input[1, 7]) AND "ROLL_IO".Input[9, 6]);
    IF #r THEN "ROLL_State".M[12, 5] := TRUE; END_IF;
    #r := "ROLL_State".M[3, 1];
    IF #r THEN "ROLL_State".M[12, 5] := FALSE; END_IF;
    // PB20, STEP 5 network 14
    #r := ((NOT "ROLL_IO".Input[9, 7]) AND ("ROLL_IO".Input[1, 6] OR "ROLL_IO".Input[1, 7]));
    IF #r THEN "ROLL_State".M[12, 6] := TRUE; END_IF;
    #r := "ROLL_State".M[3, 1];
    IF #r THEN "ROLL_State".M[12, 6] := FALSE; END_IF;
    // PB20, STEP 5 network 15
    #r := (NOT "ROLL_IO".Input[9, 6]);
    IF #r THEN "ROLL_State".M[12, 7] := TRUE; END_IF;
    #r := ("ROLL_IO".Input[9, 6] AND "ROLL_State".M[3, 1]);
    IF #r THEN "ROLL_State".M[12, 7] := FALSE; END_IF;
    // PB20, STEP 5 network 16
    #a2 := #a1;
    #a1 := "ROLL_GetDW"(DbNumber := #activeDataBlock, Index := 56);
    #r := (NOT "ROLL_IO".Input[7, 1]);
    "ROLL_TimerOp"(Number := 56, Operation := 1, Signal := #r, Preset := #a1);
    // PB20, STEP 5 network 17
    #a2 := #a1;
    #a1 := "ROLL_GetDW"(DbNumber := #activeDataBlock, Index := 65);
    #r := (NOT "ROLL_IO".Input[7, 3]);
    "ROLL_TimerOp"(Number := 65, Operation := 0, Signal := #r, Preset := #a1);
    // PB20, STEP 5 network 18
    #a2 := #a1;
    #a1 := W#16#2020;
    #r := "ROLL_IO".Input[7, 3];
    "ROLL_TimerOp"(Number := 66, Operation := 1, Signal := #r, Preset := #a1);
    // PB20, STEP 5 network 19
    #a2 := #a1;
    #a1 := "ROLL_GetDW"(DbNumber := #activeDataBlock, Index := 67);
    #r := ("ROLL_IO".Input[7, 3] AND "ROLL_State".M[150, 1]);
    "ROLL_TimerOp"(Number := 67, Operation := 0, Signal := #r, Preset := #a1);
    // PB20, STEP 5 network 20
    #a2 := #a1;
    #a1 := W#16#2005;
    #r := (NOT "ROLL_IO".Input[7, 5]);
    "ROLL_TimerOp"(Number := 96, Operation := 0, Signal := #r, Preset := #a1);
    // PB20, STEP 5 network 21
    #a2 := #a1;
    #a1 := W#16#2030;
    #r := "ROLL_IO".Input[7, 5];
    "ROLL_TimerOp"(Number := 97, Operation := 0, Signal := #r, Preset := #a1);
    // PB20, STEP 5 network 22
    #r := (((NOT "ROLL_IO".Output[18, 5]) AND "ROLL_IO".Output[18, 4]) OR ((NOT "ROLL_IO".Output[18, 7]) AND "ROLL_IO".Output[18, 6]));
    "ROLL_State".M[149, 6] := #r;
    // PB20, STEP 5 network 23
    #a2 := #a1;
    #a1 := W#16#1010;
    #r := "ROLL_State".M[148, 4];
    "ROLL_TimerOp"(Number := 89, Operation := 0, Signal := #r, Preset := #a1);
    // PB20, STEP 5 network 24
    #r := "ROLL_State".M[149, 6];
    IF #r THEN "ROLL_State".M[148, 4] := TRUE; END_IF;
    #r := "ROLL_State".S5Timers[89].Q;
    IF #r THEN "ROLL_State".M[148, 4] := FALSE; END_IF;
    // PB20, STEP 5 network 25
    #r := ("ROLL_IO".Input[8, 0] AND "ROLL_State".S5Timers[70].Q);
    "ROLL_State".M[147, 0] := #r;
    // PB20, STEP 5 network 26
    #a2 := #a1;
    #a1 := "ROLL_GetDW"(DbNumber := #activeDataBlock, Index := 75);
    #r := (NOT "ROLL_State".M[147, 0]);
    "ROLL_TimerOp"(Number := 75, Operation := 0, Signal := #r, Preset := #a1);
    // PB20, STEP 5 network 27
    #r := "ROLL_State".M[0, 3];
    "ROLL_State".M[147, 1] := #r;
    // PB20, STEP 5 network 28
    #r := ("ROLL_IO".Input[8, 2] AND "ROLL_State".S5Timers[72].Q);
    "ROLL_State".M[147, 2] := #r;
    // PB20, STEP 5 network 29
    #a2 := #a1;
    #a1 := "ROLL_GetDW"(DbNumber := #activeDataBlock, Index := 77);
    #r := (NOT "ROLL_State".M[147, 2]);
    "ROLL_TimerOp"(Number := 77, Operation := 0, Signal := #r, Preset := #a1);
    // PB20, STEP 5 network 30
    #r := "ROLL_State".M[0, 3];
    "ROLL_State".M[149, 0] := #r;
    // PB20, STEP 5 network 31
    #r := ("ROLL_State".M[147, 0] OR "ROLL_State".M[147, 2]);
    "ROLL_State".M[149, 1] := #r;
    // PB20, STEP 5 network 32
    #r := "ROLL_State".M[0, 3];
    "ROLL_State".M[149, 2] := #r;
    // PB20, STEP 5 network 33
    #r := ("ROLL_State".M[147, 0] AND "ROLL_State".M[147, 2]);
    "ROLL_State".M[149, 3] := #r;
    // PB20, STEP 5 network 34
    #r := ((NOT "ROLL_State".M[12, 6]) AND (NOT "ROLL_State".M[12, 7]) AND (NOT "ROLL_State".M[13, 4]) AND (NOT "ROLL_State".M[6, 0]) AND (NOT "ROLL_State".M[6, 2]) AND (NOT "ROLL_State".M[8, 2]) AND ("ROLL_IO".Input[1, 6] OR "ROLL_IO".Input[1, 7]) AND "ROLL_IO".Input[3, 1] AND "ROLL_IO".Input[7, 4] AND "ROLL_IO".Input[9, 6] AND "ROLL_IO".Input[9, 7] AND "ROLL_State".S5Timers[66].Q);
    "ROLL_State".M[150, 2] := #r;
    // PB20, STEP 5 network 35
    #r := ((NOT "ROLL_IO".Input[9, 2]) AND (NOT "ROLL_State".M[12, 4]) AND ("ROLL_IO".Output[18, 4] OR "ROLL_IO".Input[9, 1]) AND ("ROLL_State".M[149, 0] OR "ROLL_State".M[149, 1] OR "ROLL_State".M[149, 2] OR "ROLL_State".M[149, 3]) AND "ROLL_IO".Input[9, 0] AND "ROLL_State".M[150, 2]);
    "ROLL_IO".Output[18, 4] := #r;
    // PB20, STEP 5 network 36
    #r := ((NOT "ROLL_IO".Input[9, 2]) AND (NOT "ROLL_State".M[12, 4]) AND ("ROLL_IO".Output[18, 4] OR "ROLL_IO".Output[18, 5] OR "ROLL_IO".Input[9, 1]) AND ("ROLL_State".M[149, 2] OR "ROLL_State".M[149, 3]) AND "ROLL_IO".Input[9, 0] AND "ROLL_State".M[150, 2]);
    "ROLL_IO".Output[18, 5] := #r;
    // PB20, STEP 5 network 37
    #r := ((NOT "ROLL_IO".Input[9, 5]) AND (NOT "ROLL_State".M[12, 5]) AND ("ROLL_IO".Output[18, 6] OR "ROLL_IO".Input[9, 4]) AND ("ROLL_State".M[149, 1] OR "ROLL_State".M[149, 2] OR "ROLL_State".M[149, 3]) AND "ROLL_IO".Input[9, 3] AND "ROLL_State".M[150, 2]);
    "ROLL_IO".Output[18, 6] := #r;
    // PB20, STEP 5 network 38
    #r := ((NOT "ROLL_IO".Input[9, 5]) AND (NOT "ROLL_State".M[12, 5]) AND ("ROLL_IO".Output[18, 6] OR "ROLL_IO".Output[18, 7] OR "ROLL_IO".Input[9, 4]) AND "ROLL_IO".Input[9, 3] AND "ROLL_State".M[149, 3] AND "ROLL_State".M[150, 2]);
    "ROLL_IO".Output[18, 7] := #r;
    // PB20, STEP 5 network 39
    #r := ((NOT "ROLL_State".M[147, 0]) AND "ROLL_State".M[147, 2] AND "ROLL_State".S5Timers[75].Q);
    "ROLL_IO".Output[21, 0] := #r;
    // PB20, STEP 5 network 40
    #r := ((NOT "ROLL_State".M[147, 2]) AND "ROLL_State".M[147, 0] AND "ROLL_State".S5Timers[77].Q);
    "ROLL_IO".Output[21, 2] := #r;
    // PB20, STEP 5 network 41
    #r := "ROLL_State".M[190, 6];
    IF #r THEN "ROLL_State".M[150, 0] := TRUE; END_IF;
    #r := ((NOT "ROLL_IO".Input[0, 1]) OR (NOT "ROLL_IO".Input[7, 1]) OR (NOT "ROLL_IO".Input[7, 2]) OR (NOT "ROLL_State".M[27, 5]) OR "ROLL_IO".Input[7, 3] OR "ROLL_State".M[190, 5]);
    IF #r THEN "ROLL_State".M[150, 0] := FALSE; END_IF;
    // PB20, STEP 5 network 42
    #a2 := #a1;
    #a1 := W#16#2020;
    #r := "ROLL_IO".Input[7, 1];
    "ROLL_TimerOp"(Number := 57, Operation := 1, Signal := #r, Preset := #a1);
    // PB20, STEP 5 network 43
    #r := ((NOT "ROLL_State".M[13, 4]) AND (NOT "ROLL_State".S5Timers[61].Q) AND (((NOT "ROLL_IO".Input[7, 3]) AND "ROLL_State".S5Timers[65].Q) OR ((NOT "ROLL_State".S5Timers[67].Q) AND "ROLL_State".M[150, 1])) AND "ROLL_IO".Input[0, 2] AND "ROLL_IO".Input[3, 1] AND "ROLL_IO".Input[7, 2] AND "ROLL_State".S5Timers[57].Q);
    "ROLL_State".M[150, 1] := #r;
    // PB20, STEP 5 network 44
    #r := ("ROLL_State".M[150, 0] OR "ROLL_State".M[150, 1]);
    "ROLL_IO".Output[21, 6] := #r;
    // PB20, STEP 5 network 45
    #r := ((((NOT "ROLL_IO".Input[7, 4]) AND "ROLL_IO".Input[7, 5]) OR ((NOT "ROLL_State".S5Timers[106].Q) AND "ROLL_State".M[148, 6]) OR (NOT "ROLL_IO".Input[7, 1])) AND "ROLL_IO".Input[0, 2] AND "ROLL_IO".Input[1, 6] AND "ROLL_IO".Input[7, 0]);
    "ROLL_State".M[148, 6] := #r;
    // PB20, STEP 5 network 46
    #r := (((NOT "ROLL_State".M[151, 0]) AND (NOT "ROLL_State".M[151, 1]) AND (NOT "ROLL_State".M[151, 2]) AND (NOT "ROLL_State".M[151, 3])) OR ((NOT "ROLL_State".M[152, 3]) AND "ROLL_State".M[151, 3] AND "ROLL_State".M[153, 3] AND "ROLL_State".S5Timers[105].Q));
    IF #r THEN "ROLL_State".M[151, 0] := TRUE; END_IF;
    #r := ("ROLL_State".M[151, 1] OR "ROLL_State".M[151, 2]);
    IF #r THEN "ROLL_State".M[151, 0] := FALSE; END_IF;
    // PB20, STEP 5 network 47
    #a2 := #a1;
    #a1 := "ROLL_GetDW"(DbNumber := #activeDataBlock, Index := 102);
    #r := "ROLL_State".M[151, 0];
    "ROLL_TimerOp"(Number := 102, Operation := 0, Signal := #r, Preset := #a1);
    // PB20, STEP 5 network 48
    #r := ((NOT "ROLL_State".S5Timers[106].Q) AND "ROLL_State".M[151, 0]);
    IF #r THEN "ROLL_State".M[152, 0] := TRUE; END_IF;
    #r := ((NOT "ROLL_State".M[148, 6]) OR "ROLL_State".S5Timers[106].Q);
    IF #r THEN "ROLL_State".M[152, 0] := FALSE; END_IF;
    // PB20, STEP 5 network 49
    #r := ("ROLL_IO".Output[21, 5] AND "ROLL_State".M[152, 0]);
    IF #r THEN "ROLL_State".M[153, 0] := TRUE; END_IF;
    #r := (NOT "ROLL_State".M[151, 0]);
    IF #r THEN "ROLL_State".M[153, 0] := FALSE; END_IF;
    // PB20, STEP 5 network 50
    #r := ((NOT "ROLL_State".M[152, 0]) AND "ROLL_State".M[151, 0] AND "ROLL_State".M[153, 0] AND "ROLL_State".S5Timers[102].Q);
    IF #r THEN "ROLL_State".M[151, 1] := TRUE; END_IF;
    #r := "ROLL_State".M[151, 2];
    IF #r THEN "ROLL_State".M[151, 1] := FALSE; END_IF;
    // PB20, STEP 5 network 51
    #a2 := #a1;
    #a1 := "ROLL_GetDW"(DbNumber := #activeDataBlock, Index := 103);
    #r := "ROLL_State".M[151, 1];
    "ROLL_TimerOp"(Number := 103, Operation := 0, Signal := #r, Preset := #a1);
    // PB20, STEP 5 network 52
    #r := ((NOT "ROLL_State".S5Timers[106].Q) AND "ROLL_State".M[151, 1]);
    IF #r THEN "ROLL_State".M[152, 1] := TRUE; END_IF;
    #r := ((NOT "ROLL_State".M[148, 6]) OR "ROLL_State".S5Timers[106].Q);
    IF #r THEN "ROLL_State".M[152, 1] := FALSE; END_IF;
    // PB20, STEP 5 network 53
    #r := ("ROLL_IO".Output[20, 6] AND "ROLL_State".M[152, 1]);
    IF #r THEN "ROLL_State".M[153, 1] := TRUE; END_IF;
    #r := (NOT "ROLL_State".M[151, 1]);
    IF #r THEN "ROLL_State".M[153, 1] := FALSE; END_IF;
    // PB20, STEP 5 network 54
    #r := ((NOT "ROLL_State".M[152, 1]) AND "ROLL_State".M[151, 1] AND "ROLL_State".M[153, 1] AND "ROLL_State".S5Timers[103].Q);
    IF #r THEN "ROLL_State".M[151, 2] := TRUE; END_IF;
    #r := "ROLL_State".M[151, 3];
    IF #r THEN "ROLL_State".M[151, 2] := FALSE; END_IF;
    // PB20, STEP 5 network 55
    #a2 := #a1;
    #a1 := W#16#0002;
    #r := "ROLL_State".M[151, 2];
    "ROLL_TimerOp"(Number := 104, Operation := 0, Signal := #r, Preset := #a1);
    // PB20, STEP 5 network 56
    #r := ((NOT "ROLL_State".S5Timers[106].Q) AND "ROLL_State".M[151, 2]);
    IF #r THEN "ROLL_State".M[152, 2] := TRUE; END_IF;
    #r := ((NOT "ROLL_State".M[148, 6]) OR "ROLL_State".S5Timers[106].Q);
    IF #r THEN "ROLL_State".M[152, 2] := FALSE; END_IF;
    // PB20, STEP 5 network 57
    #r := ("ROLL_State".M[0, 4] AND "ROLL_State".M[152, 2]);
    IF #r THEN "ROLL_State".M[153, 2] := TRUE; END_IF;
    #r := (NOT "ROLL_State".M[151, 2]);
    IF #r THEN "ROLL_State".M[153, 2] := FALSE; END_IF;
    // PB20, STEP 5 network 58
    #r := ((NOT "ROLL_State".M[152, 2]) AND "ROLL_State".M[151, 2] AND "ROLL_State".M[153, 2] AND "ROLL_State".S5Timers[104].Q);
    IF #r THEN "ROLL_State".M[151, 3] := TRUE; END_IF;
    #r := "ROLL_State".M[151, 0];
    IF #r THEN "ROLL_State".M[151, 3] := FALSE; END_IF;
    // PB20, STEP 5 network 59
    #a2 := #a1;
    #a1 := W#16#0002;
    #r := "ROLL_State".M[151, 3];
    "ROLL_TimerOp"(Number := 105, Operation := 0, Signal := #r, Preset := #a1);
    // PB20, STEP 5 network 60
    #r := ((NOT "ROLL_State".S5Timers[106].Q) AND "ROLL_State".M[151, 3]);
    IF #r THEN "ROLL_State".M[152, 3] := TRUE; END_IF;
    #r := ((NOT "ROLL_State".M[148, 6]) OR "ROLL_State".S5Timers[106].Q);
    IF #r THEN "ROLL_State".M[152, 3] := FALSE; END_IF;
    // PB20, STEP 5 network 61
    #r := ("ROLL_State".M[0, 4] AND "ROLL_State".M[152, 3]);
    IF #r THEN "ROLL_State".M[153, 3] := TRUE; END_IF;
    #r := (NOT "ROLL_State".M[151, 3]);
    IF #r THEN "ROLL_State".M[153, 3] := FALSE; END_IF;
    // PB20, STEP 5 network 62
    #a2 := #a1;
    #a1 := W#16#2010;
    #r := ("ROLL_State".M[152, 0] OR "ROLL_State".M[152, 1] OR "ROLL_State".M[152, 2] OR "ROLL_State".M[152, 3]);
    "ROLL_TimerOp"(Number := 106, Operation := 0, Signal := #r, Preset := #a1);
    // PB20, STEP 5 network 63
    #r := ((NOT "ROLL_IO".Output[21, 4]) AND "ROLL_IO".Output[19, 5] AND "ROLL_State".M[152, 0]);
    "ROLL_IO".Output[21, 5] := #r;
    // PB20, STEP 5 network 64
    #r := "ROLL_State".M[152, 1];
    "ROLL_State".M[240, 0] := #r;
    // PB20, STEP 5 network 65
    #r := ((NOT "ROLL_IO".Output[21, 5]) AND "ROLL_State".M[152, 2]);
    "ROLL_State".M[240, 0] := #r;
    // PB20, STEP 5 network 66
    #r := "ROLL_State".M[152, 3];
    "ROLL_State".M[240, 0] := #r;
    // PB20, STEP 5 network 67
    #a2 := #a1;
    #a1 := "ROLL_GetDW"(DbNumber := #activeDataBlock, Index := 107);
    #r := ("ROLL_IO".Output[21, 6] AND "ROLL_IO".Input[0, 2]);
    "ROLL_TimerOp"(Number := 107, Operation := 1, Signal := #r, Preset := #a1);
    // PB20, STEP 5 network 68
    #r := ((("ROLL_IO".Output[21, 6] OR "ROLL_State".S5Timers[107].Q) AND "ROLL_IO".Input[0, 2]) OR ("ROLL_IO".Input[0, 1] AND "ROLL_State".M[190, 6] AND "ROLL_State".M[26, 6]));
    "ROLL_IO".Output[20, 5] := #r;
    // PB20, STEP 5 network 69
    RETURN;
END_FUNCTION

FUNCTION "ROLL_PB21" : Void
{ S7_Optimized_Access := 'TRUE' }
VERSION : 0.1
VAR_TEMP
    r : Bool;
    a1 : Word;
    a2 : Word;
    activeDataBlock : Int;
    comparisonResults : Array[0..0] of Bool;
END_VAR
BEGIN
    #r := FALSE;
    #a1 := W#16#0000;
    #a2 := W#16#0000;
    #activeDataBlock := 0;
    // PB21, STEP 5 network 1
    #activeDataBlock := 15;
    // PB21, STEP 5 network 2
    #r := ((NOT "ROLL_IO".Input[3, 6]) AND (NOT "ROLL_State".M[13, 1]) AND (NOT "ROLL_State".M[5, 6]));
    "ROLL_State".M[99, 7] := #r;
    // PB21, STEP 5 network 3
    #r := ((NOT "ROLL_State".M[13, 3]) AND (NOT "ROLL_State".M[16, 6]) AND (NOT "ROLL_State".M[6, 0]) AND (NOT "ROLL_State".M[6, 2]) AND "ROLL_IO".Input[3, 0] AND "ROLL_IO".Input[5, 0] AND "ROLL_IO".Input[5, 2] AND "ROLL_IO".Input[5, 4]);
    "ROLL_State".M[100, 0] := #r;
    // PB21, STEP 5 network 4
    #r := "ROLL_State".M[190, 6];
    IF #r THEN "ROLL_State".M[100, 1] := TRUE; END_IF;
    #r := (((NOT "ROLL_State".M[190, 6]) AND "ROLL_IO".Input[5, 3]) OR (NOT "ROLL_IO".Input[0, 1]) OR (NOT "ROLL_State".M[0, 3]) OR (NOT "ROLL_State".M[100, 0]) OR "ROLL_State".M[190, 5]);
    IF #r THEN "ROLL_State".M[100, 1] := FALSE; END_IF;
    // PB21, STEP 5 network 5
    #r := "ROLL_State".M[190, 6];
    IF #r THEN "ROLL_State".M[100, 2] := TRUE; END_IF;
    #r := (("ROLL_IO".Input[5, 3] AND "ROLL_IO".Input[5, 6]) OR (NOT "ROLL_IO".Input[0, 1]) OR (NOT "ROLL_State".M[0, 3]) OR (NOT "ROLL_State".M[100, 0]) OR "ROLL_State".M[190, 5]);
    IF #r THEN "ROLL_State".M[100, 2] := FALSE; END_IF;
    // PB21, STEP 5 network 6
    #r := "ROLL_State".M[190, 6];
    IF #r THEN "ROLL_State".M[100, 3] := TRUE; END_IF;
    #r := (((NOT "ROLL_IO".Input[7, 5]) AND (NOT "ROLL_State".M[190, 6])) OR (NOT "ROLL_IO".Input[0, 1]) OR (NOT "ROLL_State".M[0, 3]) OR (NOT "ROLL_State".M[100, 0]) OR "ROLL_State".M[190, 5] OR "ROLL_State".M[5, 6] OR "ROLL_State".M[8, 5]);
    IF #r THEN "ROLL_State".M[100, 3] := FALSE; END_IF;
    // PB21, STEP 5 network 7
    #r := "ROLL_State".M[190, 6];
    IF #r THEN "ROLL_State".M[100, 4] := TRUE; END_IF;
    #r := (((NOT "ROLL_State".M[100, 0]) AND (NOT "ROLL_State".M[190, 6])) OR (NOT "ROLL_IO".Input[0, 1]) OR (NOT "ROLL_State".M[0, 3]) OR (NOT "ROLL_State".M[99, 7]) OR "ROLL_State".M[190, 5]);
    IF #r THEN "ROLL_State".M[100, 4] := FALSE; END_IF;
    // PB21, STEP 5 network 8
    #r := ((NOT "ROLL_State".M[31, 5]) AND (NOT "ROLL_State".M[5, 6]) AND ((NOT "ROLL_IO".Input[5, 6]) OR (NOT "ROLL_State".S5Timers[70].Q)) AND "ROLL_IO".Input[0, 2] AND "ROLL_IO".Input[3, 1] AND "ROLL_State".M[100, 0]);
    "ROLL_State".M[100, 5] := #r;
    // PB21, STEP 5 network 9
    #r := ((("ROLL_IO".Input[7, 5] AND "ROLL_State".S5Timers[97].Q) OR (NOT "ROLL_State".S5Timers[96].Q)) AND "ROLL_State".M[0, 3] AND "ROLL_State".M[100, 5]);
    "ROLL_State".M[100, 6] := #r;
    // PB21, STEP 5 network 10
    #r := ((((NOT "ROLL_IO".Input[7, 5]) AND "ROLL_State".S5Timers[96].Q) OR (NOT "ROLL_State".S5Timers[97].Q)) AND "ROLL_State".M[0, 3] AND "ROLL_State".M[100, 5]);
    "ROLL_State".M[100, 7] := #r;
    // PB21, STEP 5 network 11
    #r := "ROLL_State".M[190, 6];
    IF #r THEN "ROLL_State".M[101, 1] := TRUE; END_IF;
    #r := (((NOT "ROLL_State".M[190, 6]) AND "ROLL_IO".Input[5, 3] AND "ROLL_IO".Input[5, 6] AND "ROLL_IO".Input[6, 0]) OR (NOT "ROLL_IO".Input[0, 1]) OR (NOT "ROLL_State".M[0, 3]) OR (NOT "ROLL_State".M[100, 0]) OR "ROLL_State".M[190, 5]);
    IF #r THEN "ROLL_State".M[101, 1] := FALSE; END_IF;
    // PB21, STEP 5 network 12
    #r := "ROLL_State".M[190, 6];
    IF #r THEN "ROLL_State".M[101, 2] := TRUE; END_IF;
    #r := (((NOT "ROLL_State".M[190, 6]) AND "ROLL_IO".Input[5, 3] AND "ROLL_IO".Input[5, 6] AND "ROLL_IO".Input[6, 0]) OR (NOT "ROLL_IO".Input[0, 1]) OR (NOT "ROLL_State".M[0, 3]) OR (NOT "ROLL_State".M[100, 0]) OR "ROLL_State".M[190, 5]);
    IF #r THEN "ROLL_State".M[101, 2] := FALSE; END_IF;
    // PB21, STEP 5 network 13
    #r := "ROLL_State".M[190, 6];
    IF #r THEN "ROLL_State".M[101, 3] := TRUE; END_IF;
    #r := (((NOT "ROLL_State".M[190, 6]) AND ((NOT "ROLL_IO".Input[7, 5]) OR "ROLL_IO".Input[6, 0])) OR (NOT "ROLL_IO".Input[0, 1]) OR (NOT "ROLL_State".M[0, 3]) OR (NOT "ROLL_State".M[100, 0]) OR "ROLL_State".M[190, 5] OR "ROLL_State".M[5, 6] OR "ROLL_State".M[8, 5]);
    IF #r THEN "ROLL_State".M[101, 3] := FALSE; END_IF;
    // PB21, STEP 5 network 14
    #r := "ROLL_State".M[190, 6];
    IF #r THEN "ROLL_State".M[101, 4] := TRUE; END_IF;
    #r := (((NOT "ROLL_State".M[190, 6]) AND "ROLL_IO".Input[6, 0]) OR (NOT "ROLL_IO".Input[0, 1]) OR (NOT "ROLL_State".M[0, 3]) OR (NOT "ROLL_State".M[100, 0]) OR (NOT "ROLL_State".M[99, 7]) OR "ROLL_State".M[190, 5]);
    IF #r THEN "ROLL_State".M[101, 4] := FALSE; END_IF;
    // PB21, STEP 5 network 15
    #a2 := #a1;
    #a1 := W#16#2005;
    #r := "ROLL_IO".Input[6, 0];
    "ROLL_TimerOp"(Number := 121, Operation := 0, Signal := #r, Preset := #a1);
    // PB21, STEP 5 network 16
    #r := ((NOT "ROLL_State".M[31, 5]) AND (NOT "ROLL_State".M[5, 6]) AND (((NOT "ROLL_State".S5Timers[121].Q) AND "ROLL_State".M[101, 5]) OR (NOT "ROLL_IO".Input[6, 0])) AND "ROLL_IO".Input[0, 2] AND "ROLL_IO".Input[3, 1] AND "ROLL_State".M[100, 0]);
    "ROLL_State".M[101, 5] := #r;
    // PB21, STEP 5 network 17
    #r := ((("ROLL_IO".Input[7, 5] AND "ROLL_State".S5Timers[97].Q) OR (NOT "ROLL_State".S5Timers[96].Q)) AND "ROLL_State".M[101, 5]);
    "ROLL_State".M[101, 6] := #r;
    // PB21, STEP 5 network 18
    #r := ((((NOT "ROLL_IO".Input[7, 5]) AND "ROLL_State".S5Timers[96].Q) OR (NOT "ROLL_State".S5Timers[97].Q)) AND "ROLL_State".M[101, 5]);
    "ROLL_State".M[101, 7] := #r;
    // PB21, STEP 5 network 19
    #r := "ROLL_State".M[190, 6];
    IF #r THEN "ROLL_State".M[102, 1] := TRUE; END_IF;
    #r := (((NOT "ROLL_State".M[190, 6]) AND "ROLL_IO".Input[5, 3] AND "ROLL_IO".Input[5, 6] AND "ROLL_IO".Input[6, 0] AND "ROLL_IO".Input[6, 2]) OR (NOT "ROLL_IO".Input[0, 1]) OR (NOT "ROLL_State".M[0, 3]) OR (NOT "ROLL_State".M[100, 0]) OR "ROLL_State".M[190, 5]);
    IF #r THEN "ROLL_State".M[102, 1] := FALSE; END_IF;
    // PB21, STEP 5 network 20
    #r := "ROLL_State".M[190, 6];
    IF #r THEN "ROLL_State".M[102, 2] := TRUE; END_IF;
    #r := (((NOT "ROLL_State".M[190, 6]) AND "ROLL_IO".Input[6, 2]) OR (NOT "ROLL_IO".Input[0, 1]) OR (NOT "ROLL_State".M[0, 3]) OR (NOT "ROLL_State".M[100, 0]) OR "ROLL_State".M[190, 5]);
    IF #r THEN "ROLL_State".M[102, 2] := FALSE; END_IF;
    // PB21, STEP 5 network 21
    #r := "ROLL_State".M[190, 6];
    IF #r THEN "ROLL_State".M[102, 3] := TRUE; END_IF;
    #r := (((NOT "ROLL_State".M[190, 6]) AND ((NOT "ROLL_IO".Input[7, 5]) OR "ROLL_IO".Input[6, 2])) OR (NOT "ROLL_IO".Input[0, 1]) OR (NOT "ROLL_State".M[0, 3]) OR (NOT "ROLL_State".M[100, 0]) OR "ROLL_State".M[190, 5] OR "ROLL_State".M[5, 6] OR "ROLL_State".M[8, 5]);
    IF #r THEN "ROLL_State".M[102, 3] := FALSE; END_IF;
    // PB21, STEP 5 network 22
    #r := "ROLL_State".M[190, 6];
    IF #r THEN "ROLL_State".M[102, 4] := TRUE; END_IF;
    #r := (((NOT "ROLL_State".M[190, 6]) AND "ROLL_IO".Input[6, 2]) OR (NOT "ROLL_IO".Input[0, 1]) OR (NOT "ROLL_State".M[0, 3]) OR (NOT "ROLL_State".M[100, 0]) OR (NOT "ROLL_State".M[99, 7]) OR "ROLL_State".M[190, 5]);
    IF #r THEN "ROLL_State".M[102, 4] := FALSE; END_IF;
    // PB21, STEP 5 network 23
    #r := ((NOT "ROLL_State".M[31, 5]) AND (NOT "ROLL_State".M[5, 6]) AND (NOT "ROLL_State".S5Timers[72].Q) AND "ROLL_IO".Input[0, 2] AND "ROLL_IO".Input[3, 1] AND "ROLL_State".M[100, 0]);
    "ROLL_State".M[102, 5] := #r;
    // PB21, STEP 5 network 24
    #r := ((("ROLL_IO".Input[7, 5] AND "ROLL_State".S5Timers[97].Q) OR (NOT "ROLL_State".S5Timers[96].Q)) AND "ROLL_State".M[0, 3] AND "ROLL_State".M[102, 5]);
    "ROLL_State".M[102, 6] := #r;
    // PB21, STEP 5 network 25
    #r := ((((NOT "ROLL_IO".Input[7, 5]) AND "ROLL_State".S5Timers[96].Q) OR (NOT "ROLL_State".S5Timers[97].Q) OR "ROLL_State".M[0, 4]) AND "ROLL_State".M[102, 5]);
    "ROLL_State".M[102, 7] := #r;
    // PB21, STEP 5 network 26
    #r := "ROLL_State".M[190, 6];
    IF #r THEN "ROLL_State".M[105, 1] := TRUE; END_IF;
    #r := (((NOT "ROLL_State".M[190, 6]) AND "ROLL_State".M[0, 4]) OR (NOT "ROLL_IO".Input[0, 1]) OR (NOT "ROLL_State".M[0, 3]) OR (NOT "ROLL_State".M[100, 0]) OR "ROLL_State".M[190, 5]);
    IF #r THEN "ROLL_State".M[105, 1] := FALSE; END_IF;
    // PB21, STEP 5 network 27
    #r := "ROLL_State".M[190, 6];
    IF #r THEN "ROLL_State".M[105, 2] := TRUE; END_IF;
    #r := ((NOT "ROLL_IO".Input[0, 1]) OR (NOT "ROLL_State".M[0, 3]) OR (NOT "ROLL_State".M[100, 0]) OR "ROLL_IO".Input[6, 2] OR "ROLL_State".M[190, 5]);
    IF #r THEN "ROLL_State".M[105, 2] := FALSE; END_IF;
    // PB21, STEP 5 network 28
    #r := "ROLL_State".M[190, 6];
    IF #r THEN "ROLL_State".M[105, 3] := TRUE; END_IF;
    #r := (((NOT "ROLL_State".M[190, 6]) AND ((NOT "ROLL_IO".Input[7, 5]) OR "ROLL_State".M[0, 4])) OR (NOT "ROLL_IO".Input[0, 1]) OR (NOT "ROLL_State".M[0, 3]) OR (NOT "ROLL_State".M[100, 0]) OR "ROLL_State".M[190, 5] OR "ROLL_State".M[5, 6] OR "ROLL_State".M[8, 5]);
    IF #r THEN "ROLL_State".M[105, 3] := FALSE; END_IF;
    // PB21, STEP 5 network 29
    #r := "ROLL_State".M[190, 6];
    IF #r THEN "ROLL_State".M[105, 4] := TRUE; END_IF;
    #r := (((NOT "ROLL_State".M[190, 6]) AND "ROLL_State".M[0, 4]) OR (NOT "ROLL_IO".Input[0, 1]) OR (NOT "ROLL_State".M[0, 3]) OR (NOT "ROLL_State".M[100, 0]) OR (NOT "ROLL_State".M[99, 7]) OR "ROLL_State".M[190, 5]);
    IF #r THEN "ROLL_State".M[105, 4] := FALSE; END_IF;
    // PB21, STEP 5 network 30
    #a2 := #a1;
    #a1 := W#16#2005;
    #r := "ROLL_State".M[0, 4];
    "ROLL_TimerOp"(Number := 120, Operation := 0, Signal := #r, Preset := #a1);
    // PB21, STEP 5 network 31
    #r := ((NOT "ROLL_State".M[31, 5]) AND (NOT "ROLL_State".M[5, 6]) AND (((NOT "ROLL_State".S5Timers[120].Q) AND "ROLL_State".M[105, 5]) OR (NOT "ROLL_State".M[0, 4])) AND "ROLL_IO".Input[0, 2] AND "ROLL_IO".Input[3, 1] AND "ROLL_State".M[100, 0]);
    "ROLL_State".M[105, 5] := #r;
    // PB21, STEP 5 network 32
    #r := ((("ROLL_IO".Input[7, 5] AND "ROLL_State".S5Timers[97].Q) OR (NOT "ROLL_State".S5Timers[96].Q)) AND "ROLL_State".M[105, 5]);
    "ROLL_State".M[105, 6] := #r;
    // PB21, STEP 5 network 33
    #r := ((((NOT "ROLL_IO".Input[7, 5]) AND "ROLL_State".S5Timers[96].Q) OR (NOT "ROLL_State".S5Timers[97].Q)) AND "ROLL_State".M[105, 5]);
    "ROLL_State".M[105, 7] := #r;
    // PB21, STEP 5 network 34
    #r := ((((NOT "ROLL_IO".Input[5, 5]) AND ("ROLL_State".M[40, 5] OR "ROLL_State".M[42, 1]) AND "ROLL_State".M[31, 5]) OR (NOT "ROLL_IO".Input[5, 6])) AND "ROLL_IO".Input[0, 2] AND "ROLL_IO".Input[3, 1] AND "ROLL_State".M[100, 0]);
    "ROLL_State".M[103, 0] := #r;
    // PB21, STEP 5 network 35
    #r := (((NOT "ROLL_IO".Input[5, 3]) OR (NOT "ROLL_IO".Input[6, 0]) OR (NOT "ROLL_State".S5Timers[121].Q)) AND "ROLL_IO".Input[3, 1] AND "ROLL_State".M[100, 0] AND "ROLL_State".M[31, 5]);
    "ROLL_State".M[103, 3] := #r;
    // PB21, STEP 5 network 36
    #r := (((NOT "ROLL_IO".Input[5, 6]) AND "ROLL_IO".Input[0, 2]) OR (("ROLL_State".M[103, 0] OR "ROLL_State".M[103, 3]) AND "ROLL_State".S5Timers[62].Q AND "ROLL_State".S5Timers[97].Q));
    "ROLL_State".M[103, 1] := #r;
    // PB21, STEP 5 network 37
    #r := ((NOT "ROLL_IO".Input[6, 2]) AND "ROLL_IO".Input[3, 1] AND "ROLL_State".M[100, 0] AND "ROLL_State".M[31, 5]);
    "ROLL_State".M[103, 4] := #r;
    // PB21, STEP 5 network 38
    #a2 := #a1;
    #a1 := W#16#1050;
    #r := ("ROLL_IO".Output[22, 3] AND "ROLL_State".M[103, 4]);
    "ROLL_TimerOp"(Number := 119, Operation := 1, Signal := #r, Preset := #a1);
    // PB21, STEP 5 network 39
    #r := (((("ROLL_State".M[103, 0] OR "ROLL_State".M[103, 3]) AND "ROLL_State".S5Timers[96].Q) OR "ROLL_State".M[103, 4] OR "ROLL_State".S5Timers[119].Q) AND "ROLL_State".S5Timers[62].Q);
    "ROLL_State".M[103, 2] := #r;
    // PB21, STEP 5 network 40
    #r := "ROLL_State".M[190, 6];
    IF #r THEN "ROLL_State".M[104, 0] := TRUE; END_IF;
    #r := (((NOT "ROLL_State".M[190, 6]) AND ((NOT "ROLL_IO".Input[5, 0]) OR (NOT "ROLL_IO".Input[5, 2]) OR (NOT "ROLL_IO".Input[5, 4]))) OR (NOT "ROLL_IO".Input[0, 1]) OR (NOT "ROLL_IO".Input[7, 0]) OR (NOT "ROLL_State".M[26, 5]) OR (NOT "ROLL_State".M[99, 7]) OR "ROLL_State".M[16, 6] OR "ROLL_State".M[190, 5]);
    IF #r THEN "ROLL_State".M[104, 0] := FALSE; END_IF;
    // PB21, STEP 5 network 41
    #r := "ROLL_State".M[190, 6];
    IF #r THEN "ROLL_State".M[104, 1] := TRUE; END_IF;
    #r := (((NOT "ROLL_State".M[190, 6]) AND ((NOT "ROLL_IO".Input[5, 0]) OR (NOT "ROLL_IO".Input[5, 2]) OR (NOT "ROLL_IO".Input[5, 4]))) OR (NOT "ROLL_IO".Input[0, 1]) OR (NOT "ROLL_State".M[26, 0]) OR (NOT "ROLL_State".M[99, 7]) OR "ROLL_State".M[16, 6] OR "ROLL_State".M[190, 5]);
    IF #r THEN "ROLL_State".M[104, 1] := FALSE; END_IF;
    // PB21, STEP 5 network 42
    #r := "ROLL_State".M[190, 6];
    IF #r THEN "ROLL_State".M[104, 4] := TRUE; END_IF;
    #r := (((NOT "ROLL_State".M[190, 6]) AND ((NOT "ROLL_IO".Input[5, 0]) OR (NOT "ROLL_IO".Input[5, 2]) OR (NOT "ROLL_IO".Input[5, 4]))) OR (NOT "ROLL_IO".Input[0, 1]) OR (NOT "ROLL_IO".Input[4, 7]) OR (NOT "ROLL_State".M[27, 4]) OR (NOT "ROLL_State".M[99, 7]) OR "ROLL_State".M[16, 6] OR "ROLL_State".M[190, 5]);
    IF #r THEN "ROLL_State".M[104, 4] := FALSE; END_IF;
    // PB21, STEP 5 network 43
    #r := "ROLL_State".M[190, 6];
    IF #r THEN "ROLL_State".M[104, 5] := TRUE; END_IF;
    #r := (((NOT "ROLL_State".M[190, 6]) AND "ROLL_IO".Input[5, 3] AND "ROLL_IO".Input[5, 6] AND "ROLL_IO".Input[6, 0] AND "ROLL_IO".Input[6, 2]) OR (NOT "ROLL_IO".Input[0, 1]) OR (NOT "ROLL_State".M[100, 0]) OR (NOT "ROLL_State".M[24, 1]) OR "ROLL_State".M[190, 5]);
    IF #r THEN "ROLL_State".M[104, 5] := FALSE; END_IF;
    // PB21, STEP 5 network 44
    #r := "ROLL_State".M[190, 6];
    IF #r THEN "ROLL_State".M[104, 6] := TRUE; END_IF;
    #r := (((NOT "ROLL_State".M[190, 6]) AND (("ROLL_IO".Input[5, 3] AND "ROLL_IO".Input[5, 6] AND "ROLL_IO".Input[6, 0]) OR (NOT "ROLL_IO".Input[7, 5]))) OR (NOT "ROLL_IO".Input[0, 1]) OR (NOT "ROLL_State".M[100, 0]) OR (NOT "ROLL_State".M[25, 0]) OR "ROLL_State".M[190, 5] OR "ROLL_State".M[5, 6] OR "ROLL_State".M[8, 5]);
    IF #r THEN "ROLL_State".M[104, 6] := FALSE; END_IF;
    // PB21, STEP 5 network 45
    #r := "ROLL_State".S5Timers[59].Q;
    "ROLL_IO".Output[17, 0] := #r;
    // PB21, STEP 5 network 46
    #r := ("ROLL_IO".Input[6, 5] AND "ROLL_State".M[100, 0]);
    "ROLL_IO".Output[17, 5] := #r;
    RETURN;
END_FUNCTION

FUNCTION "ROLL_PB23" : Void
{ S7_Optimized_Access := 'TRUE' }
VERSION : 0.1
VAR_TEMP
    r : Bool;
    a1 : Word;
    a2 : Word;
    activeDataBlock : Int;
    comparisonResults : Array[0..0] of Bool;
END_VAR
BEGIN
    #r := FALSE;
    #a1 := W#16#0000;
    #a2 := W#16#0000;
    #activeDataBlock := 0;
    // PB23, STEP 5 network 1
    #activeDataBlock := 15;
    // PB23, STEP 5 network 2
    #r := (("ROLL_State".M[40, 3] OR "ROLL_State".M[40, 4] OR "ROLL_State".M[40, 5]) AND "ROLL_State".M[111, 4]);
    "ROLL_State".M[240, 0] := #r;
    // PB23, STEP 5 network 3
    #a2 := #a1;
    #a1 := W#16#2120;
    #r := "ROLL_State".M[240, 0];
    "ROLL_TimerOp"(Number := 51, Operation := 1, Signal := #r, Preset := #a1);
    #r := "ROLL_State".S5Timers[51].Q;
    "ROLL_IO".Output[19, 0] := #r;
    // PB23, STEP 5 network 4
    #a2 := #a1;
    #a1 := W#16#1050;
    #r := ((NOT "ROLL_State".M[6, 1]) AND ("ROLL_State".M[40, 4] OR "ROLL_State".M[40, 5]) AND "ROLL_IO".Output[19, 0] AND "ROLL_State".M[240, 0] AND "ROLL_State".M[35, 2] AND "ROLL_State".S5Timers[70].Q);
    "ROLL_TimerOp"(Number := 52, Operation := 0, Signal := #r, Preset := #a1);
    #r := "ROLL_State".S5Timers[52].Q;
    "ROLL_IO".Output[19, 1] := #r;
    // PB23, STEP 5 network 5
    #r := ("ROLL_IO".Input[0, 2] AND "ROLL_IO".Input[0, 4]);
    IF #r THEN "ROLL_State".M[103, 7] := TRUE; END_IF;
    #r := (NOT "ROLL_State".S5Timers[59].Q);
    IF #r THEN "ROLL_State".M[103, 7] := FALSE; END_IF;
    // PB23, STEP 5 network 6
    #a2 := #a1;
    #a1 := W#16#3360;
    #r := "ROLL_State".S5Timers[59].Q;
    "ROLL_TimerOp"(Number := 76, Operation := 0, Signal := #r, Preset := #a1);
    // PB23, STEP 5 network 7
    #r := ((NOT "ROLL_State".M[13, 3]) AND (NOT "ROLL_State".M[5, 6]) AND (NOT "ROLL_State".M[6, 2]) AND (NOT "ROLL_State".M[6, 3]) AND (((NOT "ROLL_State".S5Timers[76].Q) AND "ROLL_IO".Input[2, 2]) OR "ROLL_State".M[103, 7] OR "ROLL_State".M[152, 0]) AND ("ROLL_IO".Input[2, 2] OR "ROLL_State".M[152, 0]) AND "ROLL_IO".Input[3, 4] AND "ROLL_IO".Input[5, 6] AND "ROLL_State".S5Timers[59].Q);
    "ROLL_IO".Output[19, 5] := #r;
    // PB23, STEP 5 network 8
    #r := ((NOT "ROLL_State".M[5, 6]) AND (NOT "ROLL_State".M[6, 1]) AND ("ROLL_IO".Input[0, 1] OR "ROLL_IO".Input[0, 2]) AND "ROLL_IO".Input[3, 1] AND "ROLL_IO".Input[3, 4] AND "ROLL_State".M[0, 3] AND "ROLL_State".M[100, 0] AND "ROLL_State".S5Timers[70].Q);
    "ROLL_State".M[240, 0] := #r;
    // PB23, STEP 5 network 9
    #r := ((NOT "ROLL_IO".Output[20, 6]) AND (NOT "ROLL_State".M[5, 6]) AND (NOT "ROLL_State".M[8, 5]) AND (NOT "ROLL_State".S5Timers[96].Q) AND (("ROLL_State".M[100, 0] AND "ROLL_State".M[103, 1]) OR "ROLL_State".M[102, 6] OR "ROLL_State".M[104, 6]));
    "ROLL_IO".Output[20, 4] := #r;
    "ROLL_IO".Output[22, 6] := #r;
    // PB23, STEP 5 network 10
    #r := ((NOT "ROLL_IO".Output[20, 1]) AND ("ROLL_State".M[104, 0] OR "ROLL_State".M[104, 1] OR "ROLL_State".M[104, 4] OR "ROLL_State".M[152, 1]) AND "ROLL_State".M[99, 7]);
    "ROLL_IO".Output[20, 6] := #r;
    // PB23, STEP 5 network 11
    #r := ("ROLL_State".M[102, 7] OR "ROLL_State".M[103, 2] OR "ROLL_State".M[104, 5]);
    "ROLL_State".M[240, 0] := #r;
    // PB23, STEP 5 network 12
    #r := ((NOT "ROLL_State".M[13, 4]) AND (NOT "ROLL_State".M[6, 0]) AND (NOT "ROLL_State".M[6, 2]) AND (NOT "ROLL_State".M[7, 7]) AND "ROLL_IO".Input[3, 1] AND "ROLL_IO".Input[5, 0] AND "ROLL_IO".Input[5, 2] AND "ROLL_IO".Input[5, 4] AND "ROLL_State".M[240, 0]);
    "ROLL_IO".Output[20, 1] := #r;
    // PB23, STEP 5 network 13
    #r := "ROLL_State".M[103, 1];
    "ROLL_IO".Output[22, 2] := #r;
    // PB23, STEP 5 network 14
    #r := ("ROLL_State".M[102, 1] OR "ROLL_State".M[102, 2] OR "ROLL_State".M[102, 3] OR "ROLL_State".M[102, 6] OR "ROLL_State".M[102, 7] OR "ROLL_State".M[103, 2]);
    "ROLL_IO".Output[22, 3] := #r;
    // PB23, STEP 5 network 15
    #r := "ROLL_State".S5Timers[85].Q;
    "ROLL_IO".Output[21, 3] := #r;
    // PB23, STEP 5 network 16
    #a2 := #a1;
    #a1 := W#16#1020;
    #r := "ROLL_IO".Output[20, 6];
    "ROLL_TimerOp"(Number := 47, Operation := 1, Signal := #r, Preset := #a1);
    // PB23, STEP 5 network 17
    #r := ((NOT "ROLL_IO".Output[21, 5]) AND (NOT "ROLL_IO".Output[22, 3]) AND (NOT "ROLL_IO".Output[22, 6]) AND (("ROLL_IO".Output[21, 4] AND "ROLL_State".S5Timers[47].Q) OR "ROLL_State".M[104, 0] OR "ROLL_State".M[152, 1]));
    "ROLL_IO".Output[21, 4] := #r;
    // PB23, STEP 5 network 18
    #r := ((NOT "ROLL_IO".Output[21, 4]) AND "ROLL_State".M[152, 0]);
    "ROLL_IO".Output[21, 5] := #r;
    // PB23, STEP 5 network 19
    RETURN;
END_FUNCTION

FUNCTION "ROLL_PB24" : Void
{ S7_Optimized_Access := 'TRUE' }
VERSION : 0.1
VAR_TEMP
    r : Bool;
    a1 : Word;
    a2 : Word;
    activeDataBlock : Int;
    comparisonResults : Array[0..0] of Bool;
END_VAR
BEGIN
    #r := FALSE;
    #a1 := W#16#0000;
    #a2 := W#16#0000;
    #activeDataBlock := 0;
    // PB24, STEP 5 network 1
    #activeDataBlock := 15;
    // PB24, STEP 5 network 2
    #r := ("ROLL_IO".Input[5, 0] AND "ROLL_State".M[13, 3] AND "ROLL_State".S5Timers[59].Q);
    "ROLL_State".M[240, 0] := #r;
    // PB24, STEP 5 network 3
    #a2 := #a1;
    #a1 := "ROLL_GetDW"(DbNumber := #activeDataBlock, Index := 54);
    #r := (NOT "ROLL_State".S5Timers[53].Q);
    "ROLL_TimerOp"(Number := 54, Operation := 0, Signal := #r, Preset := #a1);
    #a2 := #a1;
    #a1 := "ROLL_GetDW"(DbNumber := #activeDataBlock, Index := 53);
    #r := "ROLL_State".S5Timers[54].Q;
    "ROLL_TimerOp"(Number := 53, Operation := 1, Signal := #r, Preset := #a1);
    #r := "ROLL_State".M[240, 0];
    "ROLL_TimerOp"(Number := 53, Operation := 2, Signal := #r, Preset := #a1);
    #r := ((NOT "ROLL_State".M[40, 5]) AND "ROLL_State".S5Timers[53].Q);
    "ROLL_IO".Output[19, 4] := #r;
    // PB24, STEP 5 network 4
    RETURN;
END_FUNCTION

